// TIA Portal V17 export
// export: Created 2025-07-01T12:14:22.6243448Z, ExportSetting WithDefaults, DisplayName Totally Integrated Automation Portal, DisplayVersion V17, DisplayName TIA Portal Openness, DisplayVersion V17, DisplayName TIA Portal Version Control Interface, DisplayVersion V17, DisplayName SINAMICS Startdrive Advanced, DisplayVersion V17, DisplayName SINAMICS Startdrive G130, G150, S120, S150, SINAMICS MV, S210, DisplayVersion V17, DisplayName SINAMICS Startdrive G110M, G120, G120C, G120D, G120P, G115D, DisplayVersion V17, DisplayName STEP 7 Professional, DisplayVersion V17, DisplayName STEP 7 Safety, DisplayVersion V17, DisplayName WinCC Professional, DisplayVersion V17
FUNCTION_BLOCK "3PosLifter__Updated_V2_a4fa82_3a45ac7d-3c57-493c-83a9-58625a874be0 (3) - Copy_0df392"   // FB4, LAD
VERSION : 0.1
// stored: AutoNumber true, IsIECCheckEnabled false, UDAEnableTagReadback false
   VAR_INPUT
      L1S2Raise : Bool;
      iAreaClearConv : Bool;
      iAreaClearTransL2 : Bool;
      iAreaClear_TT : Bool;
      iAutoRunning : Bool;
      iErrorAck : Bool;
      iL1PalletPrsnt : Bool;
      iL1S1Raise : Bool;
      iL1S2Down : Bool;
      iL1S2DownOver : Bool;
      iL1S2Raise : Bool;
      iL2PalletPrsent : Bool;
      iL2S1Down : Bool;
      iL2S1Raise : Bool;
      iL2s2Raise : Bool;
      iLiffterAtPos1 : Bool;
      iLiffterAtPos2 : Bool;
      iLiffterAtPos3 : Bool;
      iLiffterAtPos4 : Bool;
      iLifterAt1 : Bool;
      iLifterAtPos1 : Bool;
      iLifterAtPos2 : Bool;
      iLifterAtPos3 : Bool;
      iLifterAtPos4 : Bool;
      iOTSFrmConv : Bool;
      iPalAtTT : Bool;
      iPalletAtL1 : Bool;
      iPalletAtL2 : Bool;
      iPalletAtLayre2 : Bool;
      iPalletAtTT : Bool;
      iPalletPrsntL1 : Bool;
      iRTRFrmConv : Bool;
      iRTRFrmTT : Bool;
      iRTRFrm_TT : Bool;
      iReacvAreaClr : Bool;
      iRecvAreaClear : Bool;
      iReset_fault : Bool;
      iRunOutActive : Bool;
      iRunOutCycle : Bool;
      iSstMode : Bool;
      iSstPB : Bool;
      iTransAreaClearConv : Bool;
      iTransAreaClr : Bool;
      ipalletPrsntAtTT : Bool;
   END_VAR
   VAR_OUTPUT
      qL1S1Down : Bool;
      qL1S1raise : Bool;
      qL1S2Down : Bool;
      qL1S2Raise : Bool;
      qL1TrnsfrConv : Bool;
      qL2S1raise : Bool;
      qL2S2Down : Bool;
      qL2S2Raise : Bool;
      qLiffterAtPos2 : Bool;
      qLifterAtPos1 : Bool;
      qLifterAtPos3 : Bool;
      qLifterAtPos4 : Bool;
      qLifterGotoPos1 : Bool;
      qOTSToNext : Bool;
      qOTSTo_TT : Bool;
      qOutput1 : Bool;
      qRTRToConv : Bool;
      qRTRToTT : Bool;
      qRTR_To_Conv : Bool;
   END_VAR
   VAR_IN_OUT
      IqRx_Frm_TT : Bool;
      iqRx_frm_Conv : Bool;
      iqTX_To_Conv : Bool;
      iqTX_To_TT : Bool;
      iqTx_To_ConvPos4 : Bool;
      iqTx_To_Rej : Bool;
   END_VAR
   VAR DB_SPECIFIC
      StateNo : Int;
      s100_StRunOutActive : Bool;
      s100_StRunOutActive_T1 : Bool;
      s100_StRunOutActive_T2 : Bool;
      s10_StRecovery : Bool;
      s10_StRecovery_T1 : Bool;
      s10_StRecovery_T2 : Bool;
      s10_StRecovery_T3 : Bool;
      s10_StRecovery_T4 : Bool;
      s10_StRecovery_T5 : Bool;
      s10_StRecovery_T6 : Bool;
      s10_StRecovery_T7 : Bool;
      s10_StRecovery_T8 : Bool;
      s110_InitialConvRun : Bool;
      s110_InitialConvRun_T1 : Bool;
      s120_StNextRdyInTransit : Bool;
      s120_StNextRdyInTransit_T1 : Bool;
      s120_StNextRdyInTransit_T2 : Bool;
      s130_StNextRdyInTransit_1 : Bool;
      s130_StNextRdyInTransit_1_T1 : Bool;
      s130_StNextRdyInTransit_1_T2 : Bool;
      s150_StWtLifterAtPosn1 : Bool;
      s150_StWtLifterAtPosn1_T1 : Bool;
      s15_StWtForFaultReset : Bool;
      s15_StWtForFaultReset_T1 : Bool;
      s160_StL1S2DownOver : Bool;
      s160_StL1S2DownOver_T1 : Bool;
      s170_StWtOTSFrmConv1 : Bool;
      s170_StWtOTSFrmConv1_T1 : Bool;
      s170_StWtOTSFrmConv1_T2 : Bool;
      s180_StWtRcvBegin : Bool;
      s180_StWtRcvBegin_T1 : Bool;
      s190_StWtL1RcvComplete : Bool;
      s190_StWtL1RcvComplete_T1 : Bool;
      s1_StWtResetRel : Bool;
      s1_StWtResetRel_T1 : Bool;
      s200_StWtForL1StprUp : Bool;
      s200_StWtForL1StprUp_T1 : Bool;
      s20_StWtForL1L2StoprsUp : Bool;
      s20_StWtForL1L2StoprsUp_T1 : Bool;
      s220_StWtL2S2Down : Bool;
      s220_StWtL2S2Down_T1 : Bool;
      s230_StWtL2TranBegin : Bool;
      s230_StWtL2TranBegin_T1 : Bool;
      s240_StWtL2TransComplete : Bool;
      s240_StWtL2TransComplete_T1 : Bool;
      s250_StWtDeforkDone : Bool;
      s250_StWtDeforkDone_Cond1 : Bool;
      s250_StWtDeforkDone_Cond2 : Bool;
      s250_StWtDeforkDone_T1 : Bool;
      s260_StChkRunOutActive1 : Bool;
      s260_StChkRunOutActive1_T1 : Bool;
      s260_StChkRunOutActive1_T2 : Bool;
      s270_StWtLifterAtPos4 : Bool;
      s270_StWtLifterAtPos4_T1 : Bool;
      s280_StWtRTRFrmConvPos4 : Bool;
      s280_StWtRTRFrmConvPos4_T1 : Bool;
      s285_StL1S2Down : Bool;
      s285_StL1S2Down_T1 : Bool;
      s290_StWtL1TransBeginPos4 : Bool;
      s290_StWtL1TransBeginPos4_T1 : Bool;
      s300_StWtTransDonePos4 : Bool;
      s300_StWtTransDonePos4_T1 : Bool;
      s30_StChkPalletPrsntL1L2 : Bool;
      s30_StChkPalletPrsntL1L2_T1 : Bool;
      s30_StChkPalletPrsntL1L2_T2 : Bool;
      s30_StChkPalletPrsntL1L2_T3 : Bool;
      s30_StChkPalletPrsntL1L2_T4 : Bool;
      s310_StChkPalletAtTT1 : Bool;
      s310_StChkPalletAtTT1_T1 : Bool;
      s310_StChkPalletAtTT1_T2 : Bool;
      s320_StWtLifterAtPos3 : Bool;
      s320_StWtLifterAtPos3_T1 : Bool;
      s330_StWtL2S1Down : Bool;
      s330_StWtL2S1Down_T1 : Bool;
      s340_StWtOTSFrmTT : Bool;
      s340_StWtOTSFrmTT_T1 : Bool;
      s350_StWtL2RecvingActive : Bool;
      s350_StWtL2RecvingActive_T1 : Bool;
      s360_StWtL2RcvDone : Bool;
      s360_StWtL2RcvDone_T1 : Bool;
      s370_StChkPalAtTT : Bool;
      s370_StChkPalAtTT_T1 : Bool;
      s370_StChkPalAtTT_T2 : Bool;
      s370_StChkPalAtTT_T3 : Bool;
      s380_StWtLifterAtPos2 : Bool;
      s380_StWtLifterAtPos2_T1 : Bool;
      s390_StWtRTRFrmTT : Bool;
      s390_StWtRTRFrmTT_T1 : Bool;
      s400_StWtL1S1Down1 : Bool;
      s400_StWtL1S1Down1_T1 : Bool;
      s40_StChkPalletAtTT : Bool;
      s40_StChkPalletAtTT_T1 : Bool;
      s40_StChkPalletAtTT_T2 : Bool;
      s410_StWtL1TransBegin : Bool;
      s410_StWtL1TransBegin_T1 : Bool;
      s420_StWtL1TransComplet : Bool;
      s420_StWtL1TransComplet_T1 : Bool;
      s430_StNextRdyInTransit_3 : Bool;
      s430_StNextRdyInTransit_3_T1 : Bool;
      s430_StNextRdyInTransit_3_T2 : Bool;
      s50_StWtLifterAtPos1 : Bool;
      s50_StWtLifterAtPos1_T1 : Bool;
      s60_StWtL1S2DownOver : Bool;
      s60_StWtL1S2DownOver_T1 : Bool;
      s70_StWtOTSFrmConv : Bool;
      s70_StWtOTSFrmConv_T1 : Bool;
      s80_StWtL1RecvBegin : Bool;
      s80_StWtL1RecvBegin_T1 : Bool;
      s90_StWtL1PalRcvDone : Bool;
      s90_StWtL1PalRcvDone_T1 : Bool;
      sOTSTimeout : Struct
         q : Bool;
      END_STRUCT;
      sSeq1Over : Bool;
      sSeq2Over : Bool;
      sSst : Bool;
      sSstPulse : Bool;
      sSstRise : Bool;
      sStWtResetRel : Bool;
      sStWtResetRel_T1 : Bool;
   END_VAR
   VAR_TEMP
      tOne : Bool;
   END_VAR
   VAR_TEMP   // added for the SCL form of the ladder/FBD networks
      _w1 : Bool;
   END_VAR
BEGIN

REGION Network 1
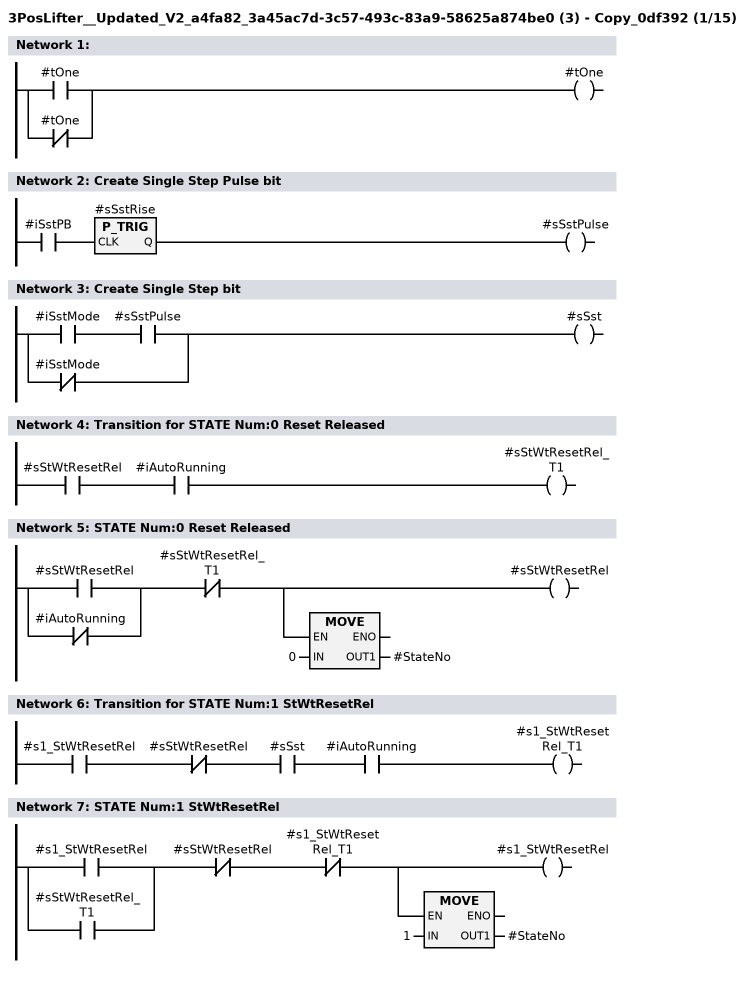
   RUNG wire#powerrail
      Contact( #tOne )
      wire#w1
      Coil( #tOne )
   END_RUNG
   RUNG wire#powerrail
      I_Contact( #tOne )
   END_RUNG wire#w1
   // the same network as SCL:
   #tOne := #tOne OR NOT #tOne;
END_REGION

REGION Network 2: Create Single Step Pulse bit
   RUNG wire#powerrail
      Contact( #iSstPB )
      P_Trig( #sSstRise )
      Coil( #sSstPulse )
   END_RUNG
   // the same network as SCL:
   #_w1 := #iSstPB AND NOT #sSstRise;   // rising edge
   #sSstRise := #iSstPB;
   #sSstPulse := #_w1;
END_REGION

REGION Network 3: Create Single Step bit
   RUNG wire#powerrail
      Contact( #iSstMode )
      Contact( #sSstPulse )
      wire#w1
      Coil( #sSst )
   END_RUNG
   RUNG wire#powerrail
      I_Contact( #iSstMode )
   END_RUNG wire#w1
   // the same network as SCL:
   #sSst := (#iSstMode AND #sSstPulse) OR NOT #iSstMode;
END_REGION

REGION Network 4: Transition for STATE Num:0 Reset Released
   RUNG wire#powerrail
      Contact( #sStWtResetRel )
      Contact( #iAutoRunning )
      Coil( #sStWtResetRel_T1 )
   END_RUNG
   // the same network as SCL:
   #sStWtResetRel_T1 := #sStWtResetRel AND #iAutoRunning;
END_REGION

REGION Network 5: STATE Num:0 Reset Released
   RUNG wire#powerrail
      Contact( #sStWtResetRel )
      wire#w1
      I_Contact( #sStWtResetRel_T1 )
      wire#w2
      Coil( #sStWtResetRel )
   END_RUNG
   RUNG wire#powerrail
      I_Contact( #iAutoRunning )
   END_RUNG wire#w1
   RUNG wire#w2
      { S7_GenerateENO := "TRUE" } Move(in := 0, out1 => #StateNo)
   END_RUNG
   // the same network as SCL:
   #sStWtResetRel := (#sStWtResetRel OR NOT #iAutoRunning) AND NOT #sStWtResetRel_T1;
   IF #sStWtResetRel THEN #StateNo := 0; END_IF;
END_REGION

REGION Network 6: Transition for STATE Num:1 StWtResetRel
   RUNG wire#powerrail
      Contact( #s1_StWtResetRel )
      I_Contact( #sStWtResetRel )
      Contact( #sSst )
      Contact( #iAutoRunning )
      Coil( #s1_StWtResetRel_T1 )
   END_RUNG
   // the same network as SCL:
   #s1_StWtResetRel_T1 := #s1_StWtResetRel AND NOT #sStWtResetRel AND #sSst AND #iAutoRunning;
END_REGION

REGION Network 7: STATE Num:1 StWtResetRel
   RUNG wire#powerrail
      Contact( #s1_StWtResetRel )
      wire#w1
      I_Contact( #sStWtResetRel )
      I_Contact( #s1_StWtResetRel_T1 )
      wire#w2
      Coil( #s1_StWtResetRel )
   END_RUNG
   RUNG wire#powerrail
      Contact( #sStWtResetRel_T1 )
   END_RUNG wire#w1
   RUNG wire#w2
      { S7_GenerateENO := "TRUE" } Move(in := 1, out1 => #StateNo)
   END_RUNG
   // the same network as SCL:
   #s1_StWtResetRel := (#s1_StWtResetRel OR #sStWtResetRel_T1) AND NOT #sStWtResetRel AND NOT #s1_StWtResetRel_T1;
   IF #s1_StWtResetRel THEN #StateNo := 1; END_IF;
END_REGION

REGION Network 8: Transition for STATE Num:10 StRecovery
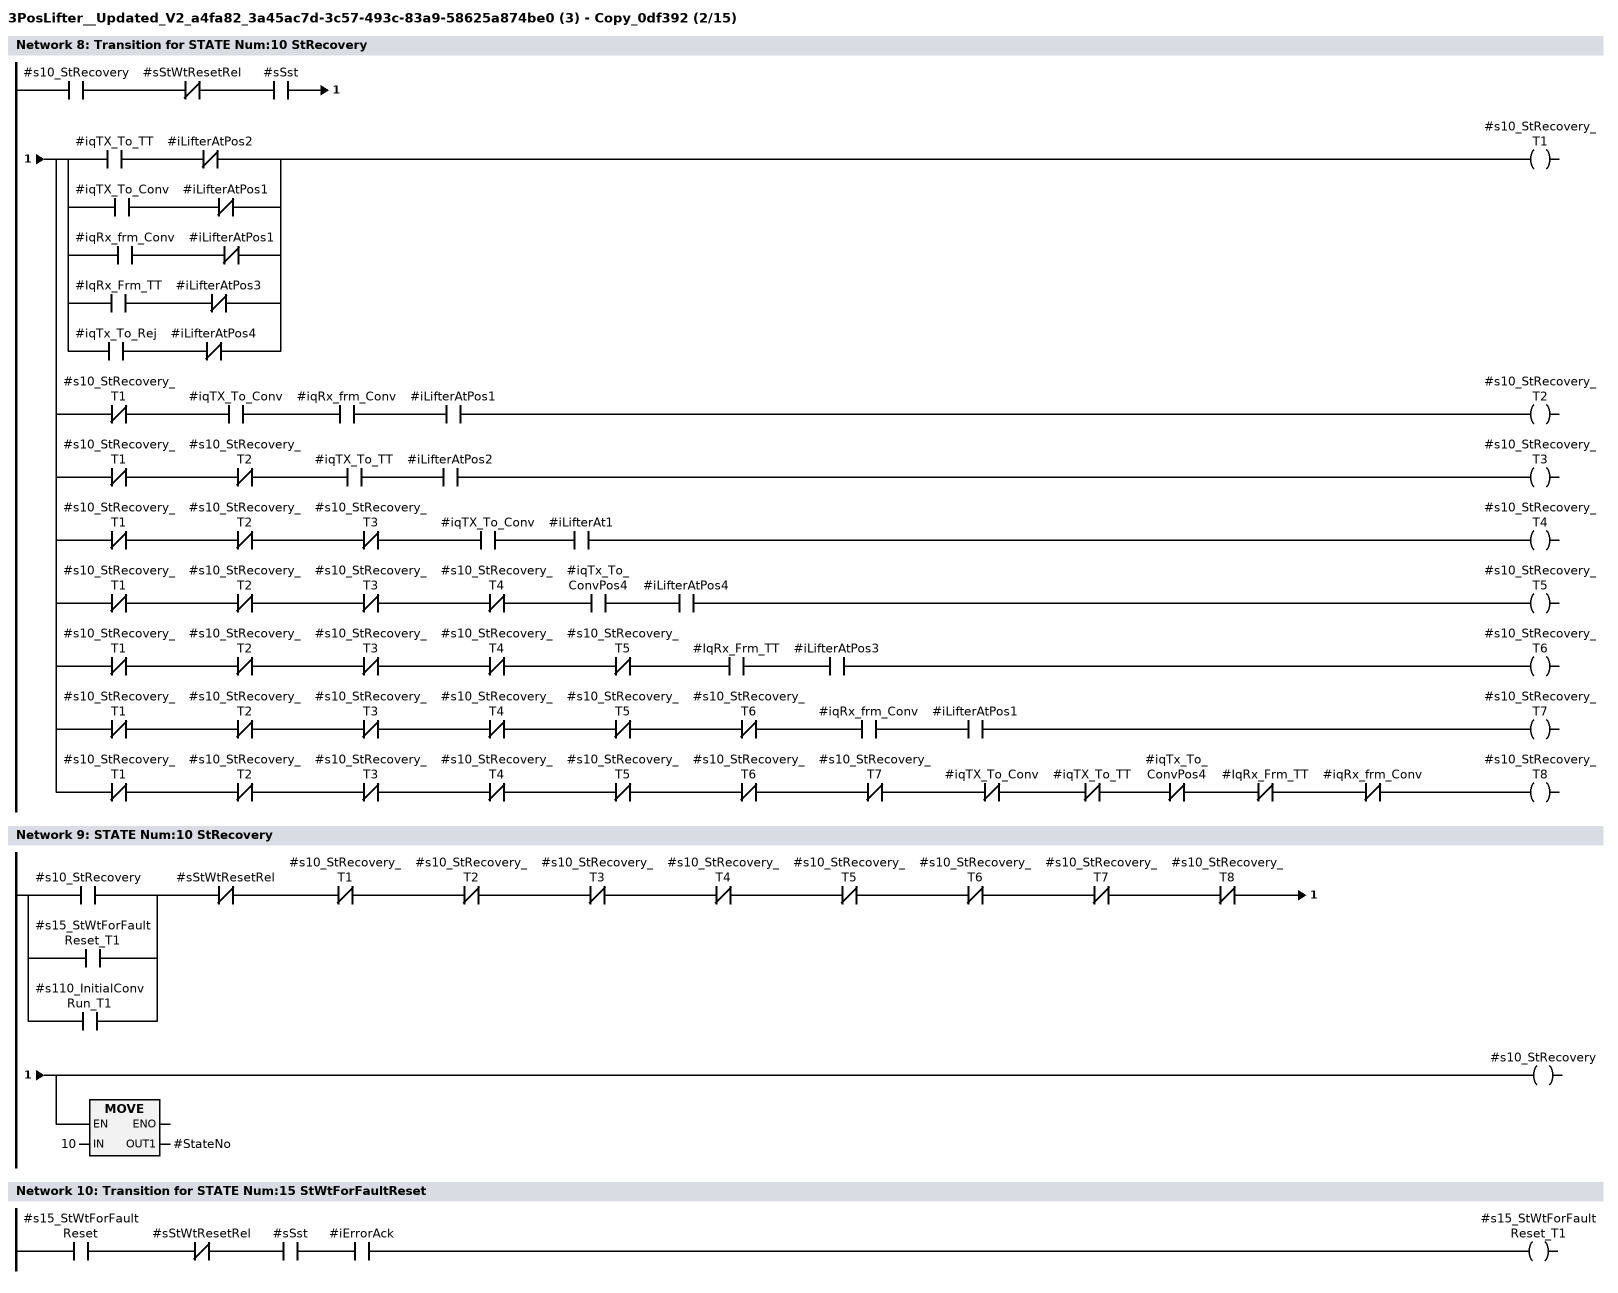
   RUNG wire#powerrail
      Contact( #s10_StRecovery )
      I_Contact( #sStWtResetRel )
      Contact( #sSst )
      wire#w1
      Contact( #iqTX_To_TT )
      I_Contact( #iLifterAtPos2 )
      wire#w2
      Coil( #s10_StRecovery_T1 )
   END_RUNG
   RUNG wire#w1
      Contact( #iqTX_To_Conv )
      I_Contact( #iLifterAtPos1 )
   END_RUNG wire#w2
   RUNG wire#w1
      Contact( #iqRx_frm_Conv )
      I_Contact( #iLifterAtPos1 )
   END_RUNG wire#w2
   RUNG wire#w1
      Contact( #IqRx_Frm_TT )
      I_Contact( #iLifterAtPos3 )
   END_RUNG wire#w2
   RUNG wire#w1
      Contact( #iqTx_To_Rej )
      I_Contact( #iLifterAtPos4 )
   END_RUNG wire#w2
   RUNG wire#w1
      I_Contact( #s10_StRecovery_T1 )
      Contact( #iqTX_To_Conv )
      Contact( #iqRx_frm_Conv )
      Contact( #iLifterAtPos1 )
      Coil( #s10_StRecovery_T2 )
   END_RUNG
   RUNG wire#w1
      I_Contact( #s10_StRecovery_T1 )
      I_Contact( #s10_StRecovery_T2 )
      Contact( #iqTX_To_TT )
      Contact( #iLifterAtPos2 )
      Coil( #s10_StRecovery_T3 )
   END_RUNG
   RUNG wire#w1
      I_Contact( #s10_StRecovery_T1 )
      I_Contact( #s10_StRecovery_T2 )
      I_Contact( #s10_StRecovery_T3 )
      Contact( #iqTX_To_Conv )
      Contact( #iLifterAt1 )
      Coil( #s10_StRecovery_T4 )
   END_RUNG
   RUNG wire#w1
      I_Contact( #s10_StRecovery_T1 )
      I_Contact( #s10_StRecovery_T2 )
      I_Contact( #s10_StRecovery_T3 )
      I_Contact( #s10_StRecovery_T4 )
      Contact( #iqTx_To_ConvPos4 )
      Contact( #iLifterAtPos4 )
      Coil( #s10_StRecovery_T5 )
   END_RUNG
   RUNG wire#w1
      I_Contact( #s10_StRecovery_T1 )
      I_Contact( #s10_StRecovery_T2 )
      I_Contact( #s10_StRecovery_T3 )
      I_Contact( #s10_StRecovery_T4 )
      I_Contact( #s10_StRecovery_T5 )
      Contact( #IqRx_Frm_TT )
      Contact( #iLifterAtPos3 )
      Coil( #s10_StRecovery_T6 )
   END_RUNG
   RUNG wire#w1
      I_Contact( #s10_StRecovery_T1 )
      I_Contact( #s10_StRecovery_T2 )
      I_Contact( #s10_StRecovery_T3 )
      I_Contact( #s10_StRecovery_T4 )
      I_Contact( #s10_StRecovery_T5 )
      I_Contact( #s10_StRecovery_T6 )
      Contact( #iqRx_frm_Conv )
      Contact( #iLifterAtPos1 )
      Coil( #s10_StRecovery_T7 )
   END_RUNG
   RUNG wire#w1
      I_Contact( #s10_StRecovery_T1 )
      I_Contact( #s10_StRecovery_T2 )
      I_Contact( #s10_StRecovery_T3 )
      I_Contact( #s10_StRecovery_T4 )
      I_Contact( #s10_StRecovery_T5 )
      I_Contact( #s10_StRecovery_T6 )
      I_Contact( #s10_StRecovery_T7 )
      I_Contact( #iqTX_To_Conv )
      I_Contact( #iqTX_To_TT )
      I_Contact( #iqTx_To_ConvPos4 )
      I_Contact( #IqRx_Frm_TT )
      I_Contact( #iqRx_frm_Conv )
      Coil( #s10_StRecovery_T8 )
   END_RUNG
   // the same network as SCL:
   #_w1 := #s10_StRecovery AND NOT #sStWtResetRel AND #sSst;
   #s10_StRecovery_T1 := #_w1 AND ((#iqTX_To_TT AND NOT #iLifterAtPos2) OR (#iqTX_To_Conv AND NOT #iLifterAtPos1) OR (#iqRx_frm_Conv AND NOT #iLifterAtPos1) OR (#IqRx_Frm_TT AND NOT #iLifterAtPos3) OR (#iqTx_To_Rej AND NOT #iLifterAtPos4));
   #s10_StRecovery_T2 := #_w1 AND NOT #s10_StRecovery_T1 AND #iqTX_To_Conv AND #iqRx_frm_Conv AND #iLifterAtPos1;
   #s10_StRecovery_T3 := #_w1 AND NOT #s10_StRecovery_T1 AND NOT #s10_StRecovery_T2 AND #iqTX_To_TT AND #iLifterAtPos2;
   #s10_StRecovery_T4 := #_w1 AND NOT #s10_StRecovery_T1 AND NOT #s10_StRecovery_T2 AND NOT #s10_StRecovery_T3 AND #iqTX_To_Conv AND #iLifterAt1;
   #s10_StRecovery_T5 := #_w1 AND NOT #s10_StRecovery_T1 AND NOT #s10_StRecovery_T2 AND NOT #s10_StRecovery_T3 AND NOT #s10_StRecovery_T4 AND #iqTx_To_ConvPos4 AND #iLifterAtPos4;
   #s10_StRecovery_T6 := #_w1 AND NOT #s10_StRecovery_T1 AND NOT #s10_StRecovery_T2 AND NOT #s10_StRecovery_T3 AND NOT #s10_StRecovery_T4 AND NOT #s10_StRecovery_T5 AND #IqRx_Frm_TT AND #iLifterAtPos3;
   #s10_StRecovery_T7 := #_w1 AND NOT #s10_StRecovery_T1 AND NOT #s10_StRecovery_T2 AND NOT #s10_StRecovery_T3 AND NOT #s10_StRecovery_T4 AND NOT #s10_StRecovery_T5 AND NOT #s10_StRecovery_T6 AND #iqRx_frm_Conv AND #iLifterAtPos1;
   #s10_StRecovery_T8 := #_w1 AND NOT #s10_StRecovery_T1 AND NOT #s10_StRecovery_T2 AND NOT #s10_StRecovery_T3 AND NOT #s10_StRecovery_T4 AND NOT #s10_StRecovery_T5 AND NOT #s10_StRecovery_T6 AND NOT #s10_StRecovery_T7 AND NOT #iqTX_To_Conv AND NOT #iqTX_To_TT AND NOT #iqTx_To_ConvPos4 AND NOT #IqRx_Frm_TT AND NOT #iqRx_frm_Conv;
END_REGION

REGION Network 9: STATE Num:10 StRecovery
   RUNG wire#powerrail
      Contact( #s10_StRecovery )
      wire#w1
      I_Contact( #sStWtResetRel )
      I_Contact( #s10_StRecovery_T1 )
      I_Contact( #s10_StRecovery_T2 )
      I_Contact( #s10_StRecovery_T3 )
      I_Contact( #s10_StRecovery_T4 )
      I_Contact( #s10_StRecovery_T5 )
      I_Contact( #s10_StRecovery_T6 )
      I_Contact( #s10_StRecovery_T7 )
      I_Contact( #s10_StRecovery_T8 )
      wire#w2
      Coil( #s10_StRecovery )
   END_RUNG
   RUNG wire#powerrail
      Contact( #s15_StWtForFaultReset_T1 )
   END_RUNG wire#w1
   RUNG wire#powerrail
      Contact( #s110_InitialConvRun_T1 )
   END_RUNG wire#w1
   RUNG wire#w2
      { S7_GenerateENO := "TRUE" } Move(in := 10, out1 => #StateNo)
   END_RUNG
   // the same network as SCL:
   #s10_StRecovery := (#s10_StRecovery OR #s15_StWtForFaultReset_T1 OR #s110_InitialConvRun_T1) AND NOT #sStWtResetRel AND NOT #s10_StRecovery_T1 AND NOT #s10_StRecovery_T2 AND NOT #s10_StRecovery_T3 AND NOT #s10_StRecovery_T4 AND NOT #s10_StRecovery_T5 AND NOT #s10_StRecovery_T6 AND NOT #s10_StRecovery_T7 AND NOT #s10_StRecovery_T8;
   IF #s10_StRecovery THEN #StateNo := 10; END_IF;
END_REGION

REGION Network 10: Transition for STATE Num:15 StWtForFaultReset
   RUNG wire#powerrail
      Contact( #s15_StWtForFaultReset )
      I_Contact( #sStWtResetRel )
      Contact( #sSst )
      Contact( #iErrorAck )
      Coil( #s15_StWtForFaultReset_T1 )
   END_RUNG
   // the same network as SCL:
   #s15_StWtForFaultReset_T1 := #s15_StWtForFaultReset AND NOT #sStWtResetRel AND #sSst AND #iErrorAck;
END_REGION

REGION Network 11: STATE Num:15 StWtForFaultReset
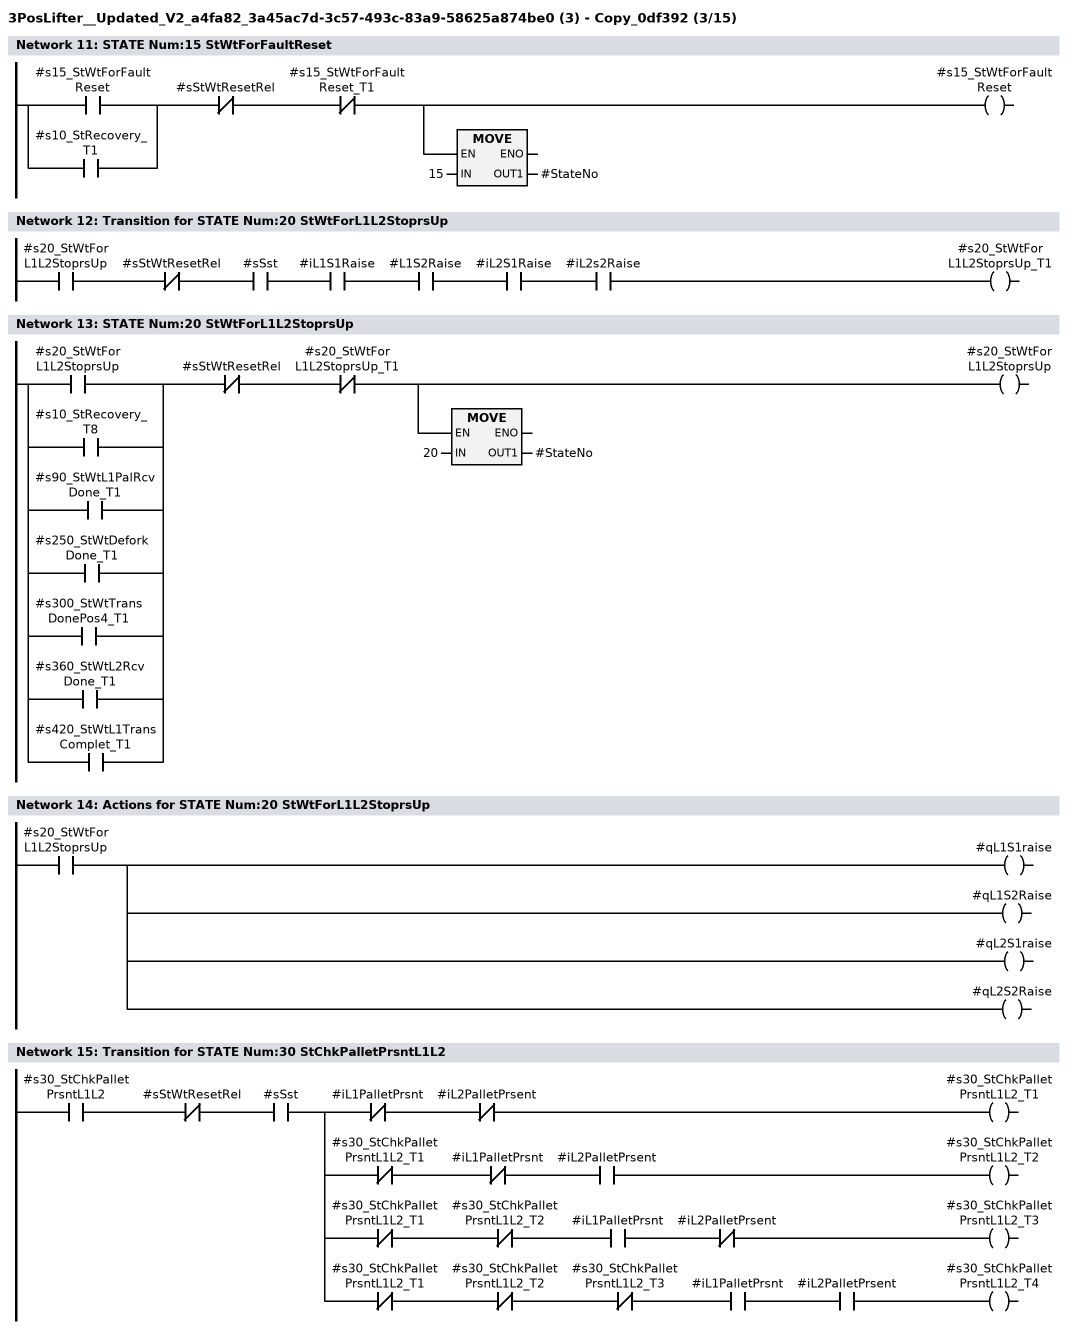
   RUNG wire#powerrail
      Contact( #s15_StWtForFaultReset )
      wire#w1
      I_Contact( #sStWtResetRel )
      I_Contact( #s15_StWtForFaultReset_T1 )
      wire#w2
      Coil( #s15_StWtForFaultReset )
   END_RUNG
   RUNG wire#powerrail
      Contact( #s10_StRecovery_T1 )
   END_RUNG wire#w1
   RUNG wire#w2
      { S7_GenerateENO := "TRUE" } Move(in := 15, out1 => #StateNo)
   END_RUNG
   // the same network as SCL:
   #s15_StWtForFaultReset := (#s15_StWtForFaultReset OR #s10_StRecovery_T1) AND NOT #sStWtResetRel AND NOT #s15_StWtForFaultReset_T1;
   IF #s15_StWtForFaultReset THEN #StateNo := 15; END_IF;
END_REGION

REGION Network 12: Transition for STATE Num:20 StWtForL1L2StoprsUp
   RUNG wire#powerrail
      Contact( #s20_StWtForL1L2StoprsUp )
      I_Contact( #sStWtResetRel )
      Contact( #sSst )
      Contact( #iL1S1Raise )
      Contact( #L1S2Raise )
      Contact( #iL2S1Raise )
      Contact( #iL2s2Raise )
      Coil( #s20_StWtForL1L2StoprsUp_T1 )
   END_RUNG
   // the same network as SCL:
   #s20_StWtForL1L2StoprsUp_T1 := #s20_StWtForL1L2StoprsUp AND NOT #sStWtResetRel AND #sSst AND #iL1S1Raise AND #L1S2Raise AND #iL2S1Raise AND #iL2s2Raise;
END_REGION

REGION Network 13: STATE Num:20 StWtForL1L2StoprsUp
   RUNG wire#powerrail
      Contact( #s20_StWtForL1L2StoprsUp )
      wire#w1
      I_Contact( #sStWtResetRel )
      I_Contact( #s20_StWtForL1L2StoprsUp_T1 )
      wire#w2
      Coil( #s20_StWtForL1L2StoprsUp )
   END_RUNG
   RUNG wire#powerrail
      Contact( #s10_StRecovery_T8 )
   END_RUNG wire#w1
   RUNG wire#powerrail
      Contact( #s90_StWtL1PalRcvDone_T1 )
   END_RUNG wire#w1
   RUNG wire#powerrail
      Contact( #s250_StWtDeforkDone_T1 )
   END_RUNG wire#w1
   RUNG wire#powerrail
      Contact( #s300_StWtTransDonePos4_T1 )
   END_RUNG wire#w1
   RUNG wire#powerrail
      Contact( #s360_StWtL2RcvDone_T1 )
   END_RUNG wire#w1
   RUNG wire#powerrail
      Contact( #s420_StWtL1TransComplet_T1 )
   END_RUNG wire#w1
   RUNG wire#w2
      { S7_GenerateENO := "TRUE" } Move(in := 20, out1 => #StateNo)
   END_RUNG
   // the same network as SCL:
   #s20_StWtForL1L2StoprsUp := (#s20_StWtForL1L2StoprsUp OR #s10_StRecovery_T8 OR #s90_StWtL1PalRcvDone_T1 OR #s250_StWtDeforkDone_T1 OR #s300_StWtTransDonePos4_T1 OR #s360_StWtL2RcvDone_T1 OR #s420_StWtL1TransComplet_T1) AND NOT #sStWtResetRel AND NOT #s20_StWtForL1L2StoprsUp_T1;
   IF #s20_StWtForL1L2StoprsUp THEN #StateNo := 20; END_IF;
END_REGION

REGION Network 14: Actions for STATE Num:20 StWtForL1L2StoprsUp
   RUNG wire#powerrail
      Contact( #s20_StWtForL1L2StoprsUp )
      wire#w1
      Coil( #qL1S1raise )
   END_RUNG
   RUNG wire#w1
      Coil( #qL1S2Raise )
   END_RUNG
   RUNG wire#w1
      Coil( #qL2S1raise )
   END_RUNG
   RUNG wire#w1
      Coil( #qL2S2Raise )
   END_RUNG
   // the same network as SCL:
   #qL1S1raise := #s20_StWtForL1L2StoprsUp;
   #qL1S2Raise := #s20_StWtForL1L2StoprsUp;
   #qL2S1raise := #s20_StWtForL1L2StoprsUp;
   #qL2S2Raise := #s20_StWtForL1L2StoprsUp;
END_REGION

REGION Network 15: Transition for STATE Num:30 StChkPalletPrsntL1L2
   RUNG wire#powerrail
      Contact( #s30_StChkPalletPrsntL1L2 )
      I_Contact( #sStWtResetRel )
      Contact( #sSst )
      wire#w1
      I_Contact( #iL1PalletPrsnt )
      I_Contact( #iL2PalletPrsent )
      Coil( #s30_StChkPalletPrsntL1L2_T1 )
   END_RUNG
   RUNG wire#w1
      I_Contact( #s30_StChkPalletPrsntL1L2_T1 )
      I_Contact( #iL1PalletPrsnt )
      Contact( #iL2PalletPrsent )
      Coil( #s30_StChkPalletPrsntL1L2_T2 )
   END_RUNG
   RUNG wire#w1
      I_Contact( #s30_StChkPalletPrsntL1L2_T1 )
      I_Contact( #s30_StChkPalletPrsntL1L2_T2 )
      Contact( #iL1PalletPrsnt )
      I_Contact( #iL2PalletPrsent )
      Coil( #s30_StChkPalletPrsntL1L2_T3 )
   END_RUNG
   RUNG wire#w1
      I_Contact( #s30_StChkPalletPrsntL1L2_T1 )
      I_Contact( #s30_StChkPalletPrsntL1L2_T2 )
      I_Contact( #s30_StChkPalletPrsntL1L2_T3 )
      Contact( #iL1PalletPrsnt )
      Contact( #iL2PalletPrsent )
      Coil( #s30_StChkPalletPrsntL1L2_T4 )
   END_RUNG
   // the same network as SCL:
   #_w1 := #s30_StChkPalletPrsntL1L2 AND NOT #sStWtResetRel AND #sSst;
   #s30_StChkPalletPrsntL1L2_T1 := #_w1 AND NOT #iL1PalletPrsnt AND NOT #iL2PalletPrsent;
   #s30_StChkPalletPrsntL1L2_T2 := #_w1 AND NOT #s30_StChkPalletPrsntL1L2_T1 AND NOT #iL1PalletPrsnt AND #iL2PalletPrsent;
   #s30_StChkPalletPrsntL1L2_T3 := #_w1 AND NOT #s30_StChkPalletPrsntL1L2_T1 AND NOT #s30_StChkPalletPrsntL1L2_T2 AND #iL1PalletPrsnt AND NOT #iL2PalletPrsent;
   #s30_StChkPalletPrsntL1L2_T4 := #_w1 AND NOT #s30_StChkPalletPrsntL1L2_T1 AND NOT #s30_StChkPalletPrsntL1L2_T2 AND NOT #s30_StChkPalletPrsntL1L2_T3 AND #iL1PalletPrsnt AND #iL2PalletPrsent;
END_REGION

REGION Network 16: STATE Num:30 StChkPalletPrsntL1L2
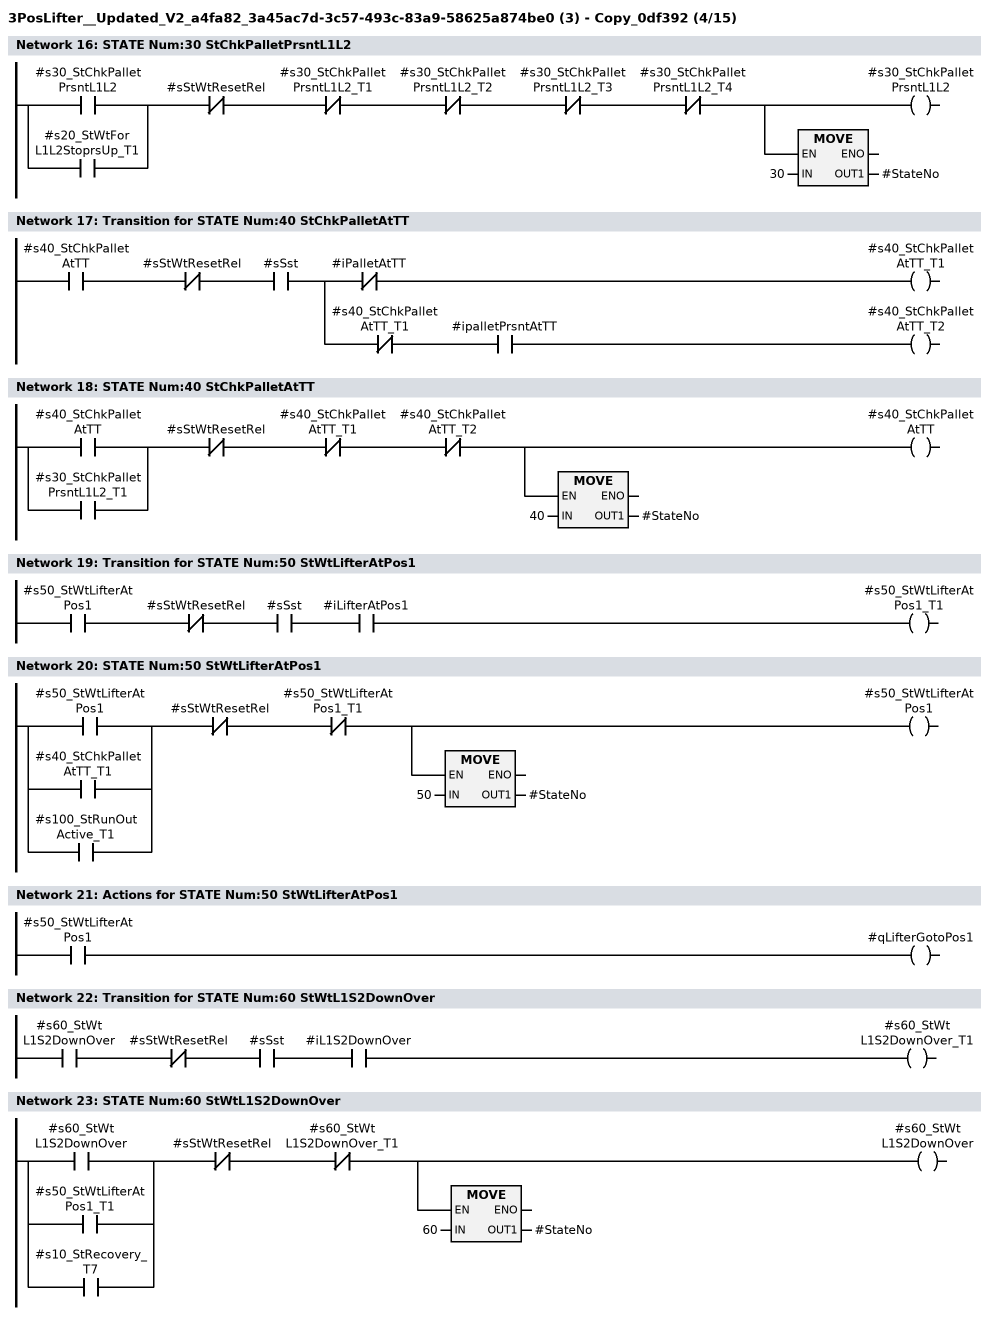
   RUNG wire#powerrail
      Contact( #s30_StChkPalletPrsntL1L2 )
      wire#w1
      I_Contact( #sStWtResetRel )
      I_Contact( #s30_StChkPalletPrsntL1L2_T1 )
      I_Contact( #s30_StChkPalletPrsntL1L2_T2 )
      I_Contact( #s30_StChkPalletPrsntL1L2_T3 )
      I_Contact( #s30_StChkPalletPrsntL1L2_T4 )
      wire#w2
      Coil( #s30_StChkPalletPrsntL1L2 )
   END_RUNG
   RUNG wire#powerrail
      Contact( #s20_StWtForL1L2StoprsUp_T1 )
   END_RUNG wire#w1
   RUNG wire#w2
      { S7_GenerateENO := "TRUE" } Move(in := 30, out1 => #StateNo)
   END_RUNG
   // the same network as SCL:
   #s30_StChkPalletPrsntL1L2 := (#s30_StChkPalletPrsntL1L2 OR #s20_StWtForL1L2StoprsUp_T1) AND NOT #sStWtResetRel AND NOT #s30_StChkPalletPrsntL1L2_T1 AND NOT #s30_StChkPalletPrsntL1L2_T2 AND NOT #s30_StChkPalletPrsntL1L2_T3 AND NOT #s30_StChkPalletPrsntL1L2_T4;
   IF #s30_StChkPalletPrsntL1L2 THEN #StateNo := 30; END_IF;
END_REGION

REGION Network 17: Transition for STATE Num:40 StChkPalletAtTT
   RUNG wire#powerrail
      Contact( #s40_StChkPalletAtTT )
      I_Contact( #sStWtResetRel )
      Contact( #sSst )
      wire#w1
      I_Contact( #iPalletAtTT )
      Coil( #s40_StChkPalletAtTT_T1 )
   END_RUNG
   RUNG wire#w1
      I_Contact( #s40_StChkPalletAtTT_T1 )
      Contact( #ipalletPrsntAtTT )
      Coil( #s40_StChkPalletAtTT_T2 )
   END_RUNG
   // the same network as SCL:
   #_w1 := #s40_StChkPalletAtTT AND NOT #sStWtResetRel AND #sSst;
   #s40_StChkPalletAtTT_T1 := #_w1 AND NOT #iPalletAtTT;
   #s40_StChkPalletAtTT_T2 := #_w1 AND NOT #s40_StChkPalletAtTT_T1 AND #ipalletPrsntAtTT;
END_REGION

REGION Network 18: STATE Num:40 StChkPalletAtTT
   RUNG wire#powerrail
      Contact( #s40_StChkPalletAtTT )
      wire#w1
      I_Contact( #sStWtResetRel )
      I_Contact( #s40_StChkPalletAtTT_T1 )
      I_Contact( #s40_StChkPalletAtTT_T2 )
      wire#w2
      Coil( #s40_StChkPalletAtTT )
   END_RUNG
   RUNG wire#powerrail
      Contact( #s30_StChkPalletPrsntL1L2_T1 )
   END_RUNG wire#w1
   RUNG wire#w2
      { S7_GenerateENO := "TRUE" } Move(in := 40, out1 => #StateNo)
   END_RUNG
   // the same network as SCL:
   #s40_StChkPalletAtTT := (#s40_StChkPalletAtTT OR #s30_StChkPalletPrsntL1L2_T1) AND NOT #sStWtResetRel AND NOT #s40_StChkPalletAtTT_T1 AND NOT #s40_StChkPalletAtTT_T2;
   IF #s40_StChkPalletAtTT THEN #StateNo := 40; END_IF;
END_REGION

REGION Network 19: Transition for STATE Num:50 StWtLifterAtPos1
   RUNG wire#powerrail
      Contact( #s50_StWtLifterAtPos1 )
      I_Contact( #sStWtResetRel )
      Contact( #sSst )
      Contact( #iLifterAtPos1 )
      Coil( #s50_StWtLifterAtPos1_T1 )
   END_RUNG
   // the same network as SCL:
   #s50_StWtLifterAtPos1_T1 := #s50_StWtLifterAtPos1 AND NOT #sStWtResetRel AND #sSst AND #iLifterAtPos1;
END_REGION

REGION Network 20: STATE Num:50 StWtLifterAtPos1
   RUNG wire#powerrail
      Contact( #s50_StWtLifterAtPos1 )
      wire#w1
      I_Contact( #sStWtResetRel )
      I_Contact( #s50_StWtLifterAtPos1_T1 )
      wire#w2
      Coil( #s50_StWtLifterAtPos1 )
   END_RUNG
   RUNG wire#powerrail
      Contact( #s40_StChkPalletAtTT_T1 )
   END_RUNG wire#w1
   RUNG wire#powerrail
      Contact( #s100_StRunOutActive_T1 )
   END_RUNG wire#w1
   RUNG wire#w2
      { S7_GenerateENO := "TRUE" } Move(in := 50, out1 => #StateNo)
   END_RUNG
   // the same network as SCL:
   #s50_StWtLifterAtPos1 := (#s50_StWtLifterAtPos1 OR #s40_StChkPalletAtTT_T1 OR #s100_StRunOutActive_T1) AND NOT #sStWtResetRel AND NOT #s50_StWtLifterAtPos1_T1;
   IF #s50_StWtLifterAtPos1 THEN #StateNo := 50; END_IF;
END_REGION

REGION Network 21: Actions for STATE Num:50 StWtLifterAtPos1
   RUNG wire#powerrail
      Contact( #s50_StWtLifterAtPos1 )
      Coil( #qLifterGotoPos1 )
   END_RUNG
   // the same network as SCL:
   #qLifterGotoPos1 := #s50_StWtLifterAtPos1;
END_REGION

REGION Network 22: Transition for STATE Num:60 StWtL1S2DownOver
   RUNG wire#powerrail
      Contact( #s60_StWtL1S2DownOver )
      I_Contact( #sStWtResetRel )
      Contact( #sSst )
      Contact( #iL1S2DownOver )
      Coil( #s60_StWtL1S2DownOver_T1 )
   END_RUNG
   // the same network as SCL:
   #s60_StWtL1S2DownOver_T1 := #s60_StWtL1S2DownOver AND NOT #sStWtResetRel AND #sSst AND #iL1S2DownOver;
END_REGION

REGION Network 23: STATE Num:60 StWtL1S2DownOver
   RUNG wire#powerrail
      Contact( #s60_StWtL1S2DownOver )
      wire#w1
      I_Contact( #sStWtResetRel )
      I_Contact( #s60_StWtL1S2DownOver_T1 )
      wire#w2
      Coil( #s60_StWtL1S2DownOver )
   END_RUNG
   RUNG wire#powerrail
      Contact( #s50_StWtLifterAtPos1_T1 )
   END_RUNG wire#w1
   RUNG wire#powerrail
      Contact( #s10_StRecovery_T7 )
   END_RUNG wire#w1
   RUNG wire#w2
      { S7_GenerateENO := "TRUE" } Move(in := 60, out1 => #StateNo)
   END_RUNG
   // the same network as SCL:
   #s60_StWtL1S2DownOver := (#s60_StWtL1S2DownOver OR #s50_StWtLifterAtPos1_T1 OR #s10_StRecovery_T7) AND NOT #sStWtResetRel AND NOT #s60_StWtL1S2DownOver_T1;
   IF #s60_StWtL1S2DownOver THEN #StateNo := 60; END_IF;
END_REGION

REGION Network 24: Actions for STATE Num:60 StWtL1S2DownOver
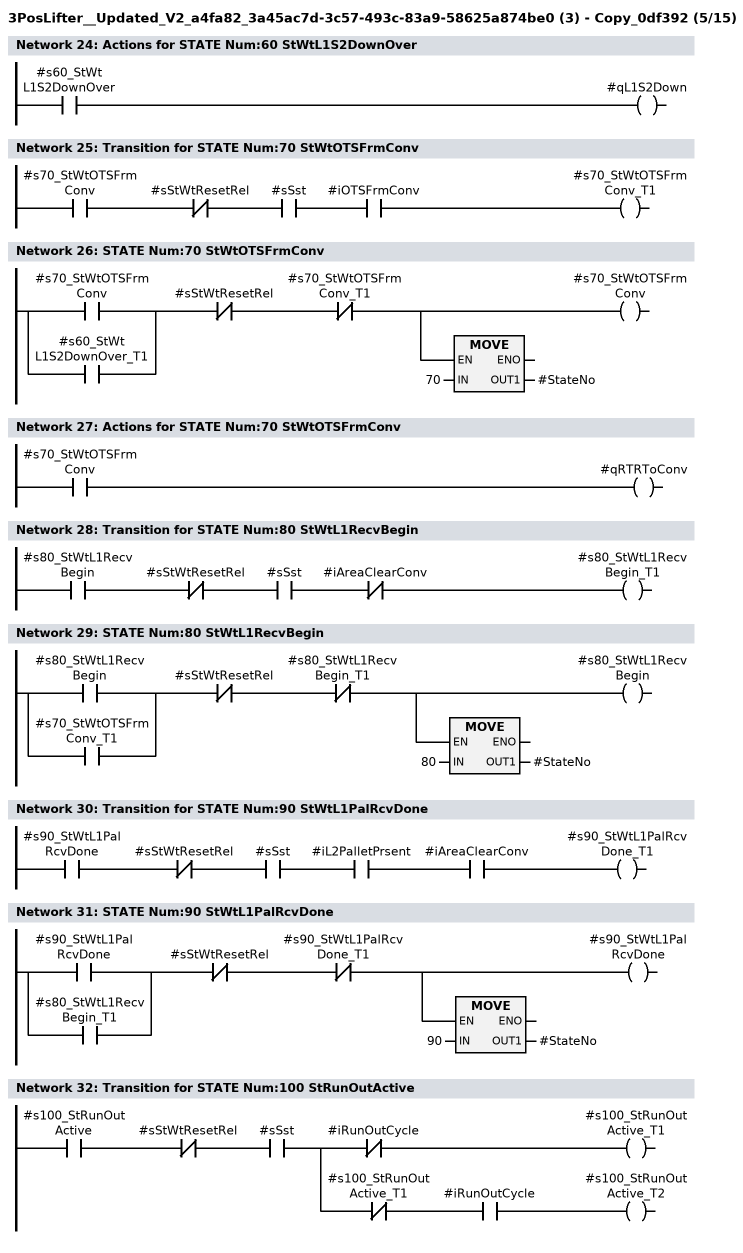
   RUNG wire#powerrail
      Contact( #s60_StWtL1S2DownOver )
      Coil( #qL1S2Down )
   END_RUNG
   // the same network as SCL:
   #qL1S2Down := #s60_StWtL1S2DownOver;
END_REGION

REGION Network 25: Transition for STATE Num:70 StWtOTSFrmConv
   RUNG wire#powerrail
      Contact( #s70_StWtOTSFrmConv )
      I_Contact( #sStWtResetRel )
      Contact( #sSst )
      Contact( #iOTSFrmConv )
      Coil( #s70_StWtOTSFrmConv_T1 )
   END_RUNG
   // the same network as SCL:
   #s70_StWtOTSFrmConv_T1 := #s70_StWtOTSFrmConv AND NOT #sStWtResetRel AND #sSst AND #iOTSFrmConv;
END_REGION

REGION Network 26: STATE Num:70 StWtOTSFrmConv
   RUNG wire#powerrail
      Contact( #s70_StWtOTSFrmConv )
      wire#w1
      I_Contact( #sStWtResetRel )
      I_Contact( #s70_StWtOTSFrmConv_T1 )
      wire#w2
      Coil( #s70_StWtOTSFrmConv )
   END_RUNG
   RUNG wire#powerrail
      Contact( #s60_StWtL1S2DownOver_T1 )
   END_RUNG wire#w1
   RUNG wire#w2
      { S7_GenerateENO := "TRUE" } Move(in := 70, out1 => #StateNo)
   END_RUNG
   // the same network as SCL:
   #s70_StWtOTSFrmConv := (#s70_StWtOTSFrmConv OR #s60_StWtL1S2DownOver_T1) AND NOT #sStWtResetRel AND NOT #s70_StWtOTSFrmConv_T1;
   IF #s70_StWtOTSFrmConv THEN #StateNo := 70; END_IF;
END_REGION

REGION Network 27: Actions for STATE Num:70 StWtOTSFrmConv
   RUNG wire#powerrail
      Contact( #s70_StWtOTSFrmConv )
      Coil( #qRTRToConv )
   END_RUNG
   // the same network as SCL:
   #qRTRToConv := #s70_StWtOTSFrmConv;
END_REGION

REGION Network 28: Transition for STATE Num:80 StWtL1RecvBegin
   RUNG wire#powerrail
      Contact( #s80_StWtL1RecvBegin )
      I_Contact( #sStWtResetRel )
      Contact( #sSst )
      I_Contact( #iAreaClearConv )
      Coil( #s80_StWtL1RecvBegin_T1 )
   END_RUNG
   // the same network as SCL:
   #s80_StWtL1RecvBegin_T1 := #s80_StWtL1RecvBegin AND NOT #sStWtResetRel AND #sSst AND NOT #iAreaClearConv;
END_REGION

REGION Network 29: STATE Num:80 StWtL1RecvBegin
   RUNG wire#powerrail
      Contact( #s80_StWtL1RecvBegin )
      wire#w1
      I_Contact( #sStWtResetRel )
      I_Contact( #s80_StWtL1RecvBegin_T1 )
      wire#w2
      Coil( #s80_StWtL1RecvBegin )
   END_RUNG
   RUNG wire#powerrail
      Contact( #s70_StWtOTSFrmConv_T1 )
   END_RUNG wire#w1
   RUNG wire#w2
      { S7_GenerateENO := "TRUE" } Move(in := 80, out1 => #StateNo)
   END_RUNG
   // the same network as SCL:
   #s80_StWtL1RecvBegin := (#s80_StWtL1RecvBegin OR #s70_StWtOTSFrmConv_T1) AND NOT #sStWtResetRel AND NOT #s80_StWtL1RecvBegin_T1;
   IF #s80_StWtL1RecvBegin THEN #StateNo := 80; END_IF;
END_REGION

REGION Network 30: Transition for STATE Num:90 StWtL1PalRcvDone
   RUNG wire#powerrail
      Contact( #s90_StWtL1PalRcvDone )
      I_Contact( #sStWtResetRel )
      Contact( #sSst )
      Contact( #iL2PalletPrsent )
      Contact( #iAreaClearConv )
      Coil( #s90_StWtL1PalRcvDone_T1 )
   END_RUNG
   // the same network as SCL:
   #s90_StWtL1PalRcvDone_T1 := #s90_StWtL1PalRcvDone AND NOT #sStWtResetRel AND #sSst AND #iL2PalletPrsent AND #iAreaClearConv;
END_REGION

REGION Network 31: STATE Num:90 StWtL1PalRcvDone
   RUNG wire#powerrail
      Contact( #s90_StWtL1PalRcvDone )
      wire#w1
      I_Contact( #sStWtResetRel )
      I_Contact( #s90_StWtL1PalRcvDone_T1 )
      wire#w2
      Coil( #s90_StWtL1PalRcvDone )
   END_RUNG
   RUNG wire#powerrail
      Contact( #s80_StWtL1RecvBegin_T1 )
   END_RUNG wire#w1
   RUNG wire#w2
      { S7_GenerateENO := "TRUE" } Move(in := 90, out1 => #StateNo)
   END_RUNG
   // the same network as SCL:
   #s90_StWtL1PalRcvDone := (#s90_StWtL1PalRcvDone OR #s80_StWtL1RecvBegin_T1) AND NOT #sStWtResetRel AND NOT #s90_StWtL1PalRcvDone_T1;
   IF #s90_StWtL1PalRcvDone THEN #StateNo := 90; END_IF;
END_REGION

REGION Network 32: Transition for STATE Num:100 StRunOutActive
   RUNG wire#powerrail
      Contact( #s100_StRunOutActive )
      I_Contact( #sStWtResetRel )
      Contact( #sSst )
      wire#w1
      I_Contact( #iRunOutCycle )
      Coil( #s100_StRunOutActive_T1 )
   END_RUNG
   RUNG wire#w1
      I_Contact( #s100_StRunOutActive_T1 )
      Contact( #iRunOutCycle )
      Coil( #s100_StRunOutActive_T2 )
   END_RUNG
   // the same network as SCL:
   #_w1 := #s100_StRunOutActive AND NOT #sStWtResetRel AND #sSst;
   #s100_StRunOutActive_T1 := #_w1 AND NOT #iRunOutCycle;
   #s100_StRunOutActive_T2 := #_w1 AND NOT #s100_StRunOutActive_T1 AND #iRunOutCycle;
END_REGION

REGION Network 33: STATE Num:100 StRunOutActive
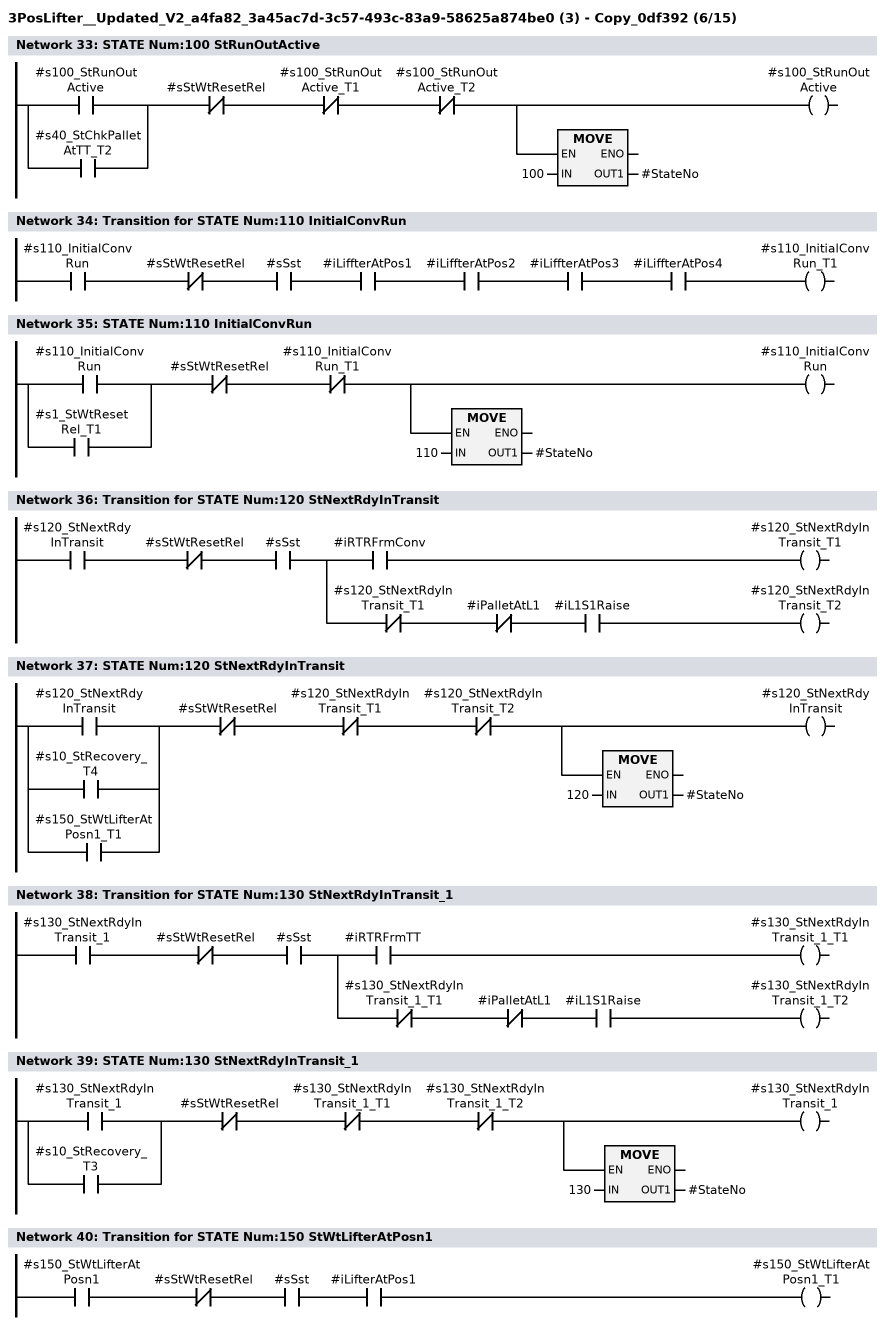
   RUNG wire#powerrail
      Contact( #s100_StRunOutActive )
      wire#w1
      I_Contact( #sStWtResetRel )
      I_Contact( #s100_StRunOutActive_T1 )
      I_Contact( #s100_StRunOutActive_T2 )
      wire#w2
      Coil( #s100_StRunOutActive )
   END_RUNG
   RUNG wire#powerrail
      Contact( #s40_StChkPalletAtTT_T2 )
   END_RUNG wire#w1
   RUNG wire#w2
      { S7_GenerateENO := "TRUE" } Move(in := 100, out1 => #StateNo)
   END_RUNG
   // the same network as SCL:
   #s100_StRunOutActive := (#s100_StRunOutActive OR #s40_StChkPalletAtTT_T2) AND NOT #sStWtResetRel AND NOT #s100_StRunOutActive_T1 AND NOT #s100_StRunOutActive_T2;
   IF #s100_StRunOutActive THEN #StateNo := 100; END_IF;
END_REGION

REGION Network 34: Transition for STATE Num:110 InitialConvRun
   RUNG wire#powerrail
      Contact( #s110_InitialConvRun )
      I_Contact( #sStWtResetRel )
      Contact( #sSst )
      Contact( #iLiffterAtPos1 )
      Contact( #iLiffterAtPos2 )
      Contact( #iLiffterAtPos3 )
      Contact( #iLiffterAtPos4 )
      Coil( #s110_InitialConvRun_T1 )
   END_RUNG
   // the same network as SCL:
   #s110_InitialConvRun_T1 := #s110_InitialConvRun AND NOT #sStWtResetRel AND #sSst AND #iLiffterAtPos1 AND #iLiffterAtPos2 AND #iLiffterAtPos3 AND #iLiffterAtPos4;
END_REGION

REGION Network 35: STATE Num:110 InitialConvRun
   RUNG wire#powerrail
      Contact( #s110_InitialConvRun )
      wire#w1
      I_Contact( #sStWtResetRel )
      I_Contact( #s110_InitialConvRun_T1 )
      wire#w2
      Coil( #s110_InitialConvRun )
   END_RUNG
   RUNG wire#powerrail
      Contact( #s1_StWtResetRel_T1 )
   END_RUNG wire#w1
   RUNG wire#w2
      { S7_GenerateENO := "TRUE" } Move(in := 110, out1 => #StateNo)
   END_RUNG
   // the same network as SCL:
   #s110_InitialConvRun := (#s110_InitialConvRun OR #s1_StWtResetRel_T1) AND NOT #sStWtResetRel AND NOT #s110_InitialConvRun_T1;
   IF #s110_InitialConvRun THEN #StateNo := 110; END_IF;
END_REGION

REGION Network 36: Transition for STATE Num:120 StNextRdyInTransit
   RUNG wire#powerrail
      Contact( #s120_StNextRdyInTransit )
      I_Contact( #sStWtResetRel )
      Contact( #sSst )
      wire#w1
      Contact( #iRTRFrmConv )
      Coil( #s120_StNextRdyInTransit_T1 )
   END_RUNG
   RUNG wire#w1
      I_Contact( #s120_StNextRdyInTransit_T1 )
      I_Contact( #iPalletAtL1 )
      Contact( #iL1S1Raise )
      Coil( #s120_StNextRdyInTransit_T2 )
   END_RUNG
   // the same network as SCL:
   #_w1 := #s120_StNextRdyInTransit AND NOT #sStWtResetRel AND #sSst;
   #s120_StNextRdyInTransit_T1 := #_w1 AND #iRTRFrmConv;
   #s120_StNextRdyInTransit_T2 := #_w1 AND NOT #s120_StNextRdyInTransit_T1 AND NOT #iPalletAtL1 AND #iL1S1Raise;
END_REGION

REGION Network 37: STATE Num:120 StNextRdyInTransit
   RUNG wire#powerrail
      Contact( #s120_StNextRdyInTransit )
      wire#w1
      I_Contact( #sStWtResetRel )
      I_Contact( #s120_StNextRdyInTransit_T1 )
      I_Contact( #s120_StNextRdyInTransit_T2 )
      wire#w2
      Coil( #s120_StNextRdyInTransit )
   END_RUNG
   RUNG wire#powerrail
      Contact( #s10_StRecovery_T4 )
   END_RUNG wire#w1
   RUNG wire#powerrail
      Contact( #s150_StWtLifterAtPosn1_T1 )
   END_RUNG wire#w1
   RUNG wire#w2
      { S7_GenerateENO := "TRUE" } Move(in := 120, out1 => #StateNo)
   END_RUNG
   // the same network as SCL:
   #s120_StNextRdyInTransit := (#s120_StNextRdyInTransit OR #s10_StRecovery_T4 OR #s150_StWtLifterAtPosn1_T1) AND NOT #sStWtResetRel AND NOT #s120_StNextRdyInTransit_T1 AND NOT #s120_StNextRdyInTransit_T2;
   IF #s120_StNextRdyInTransit THEN #StateNo := 120; END_IF;
END_REGION

REGION Network 38: Transition for STATE Num:130 StNextRdyInTransit_1
   RUNG wire#powerrail
      Contact( #s130_StNextRdyInTransit_1 )
      I_Contact( #sStWtResetRel )
      Contact( #sSst )
      wire#w1
      Contact( #iRTRFrmTT )
      Coil( #s130_StNextRdyInTransit_1_T1 )
   END_RUNG
   RUNG wire#w1
      I_Contact( #s130_StNextRdyInTransit_1_T1 )
      I_Contact( #iPalletAtL1 )
      Contact( #iL1S1Raise )
      Coil( #s130_StNextRdyInTransit_1_T2 )
   END_RUNG
   // the same network as SCL:
   #_w1 := #s130_StNextRdyInTransit_1 AND NOT #sStWtResetRel AND #sSst;
   #s130_StNextRdyInTransit_1_T1 := #_w1 AND #iRTRFrmTT;
   #s130_StNextRdyInTransit_1_T2 := #_w1 AND NOT #s130_StNextRdyInTransit_1_T1 AND NOT #iPalletAtL1 AND #iL1S1Raise;
END_REGION

REGION Network 39: STATE Num:130 StNextRdyInTransit_1
   RUNG wire#powerrail
      Contact( #s130_StNextRdyInTransit_1 )
      wire#w1
      I_Contact( #sStWtResetRel )
      I_Contact( #s130_StNextRdyInTransit_1_T1 )
      I_Contact( #s130_StNextRdyInTransit_1_T2 )
      wire#w2
      Coil( #s130_StNextRdyInTransit_1 )
   END_RUNG
   RUNG wire#powerrail
      Contact( #s10_StRecovery_T3 )
   END_RUNG wire#w1
   RUNG wire#w2
      { S7_GenerateENO := "TRUE" } Move(in := 130, out1 => #StateNo)
   END_RUNG
   // the same network as SCL:
   #s130_StNextRdyInTransit_1 := (#s130_StNextRdyInTransit_1 OR #s10_StRecovery_T3) AND NOT #sStWtResetRel AND NOT #s130_StNextRdyInTransit_1_T1 AND NOT #s130_StNextRdyInTransit_1_T2;
   IF #s130_StNextRdyInTransit_1 THEN #StateNo := 130; END_IF;
END_REGION

REGION Network 40: Transition for STATE Num:150 StWtLifterAtPosn1
   RUNG wire#powerrail
      Contact( #s150_StWtLifterAtPosn1 )
      I_Contact( #sStWtResetRel )
      Contact( #sSst )
      Contact( #iLifterAtPos1 )
      Coil( #s150_StWtLifterAtPosn1_T1 )
   END_RUNG
   // the same network as SCL:
   #s150_StWtLifterAtPosn1_T1 := #s150_StWtLifterAtPosn1 AND NOT #sStWtResetRel AND #sSst AND #iLifterAtPos1;
END_REGION

REGION Network 41: STATE Num:150 StWtLifterAtPosn1
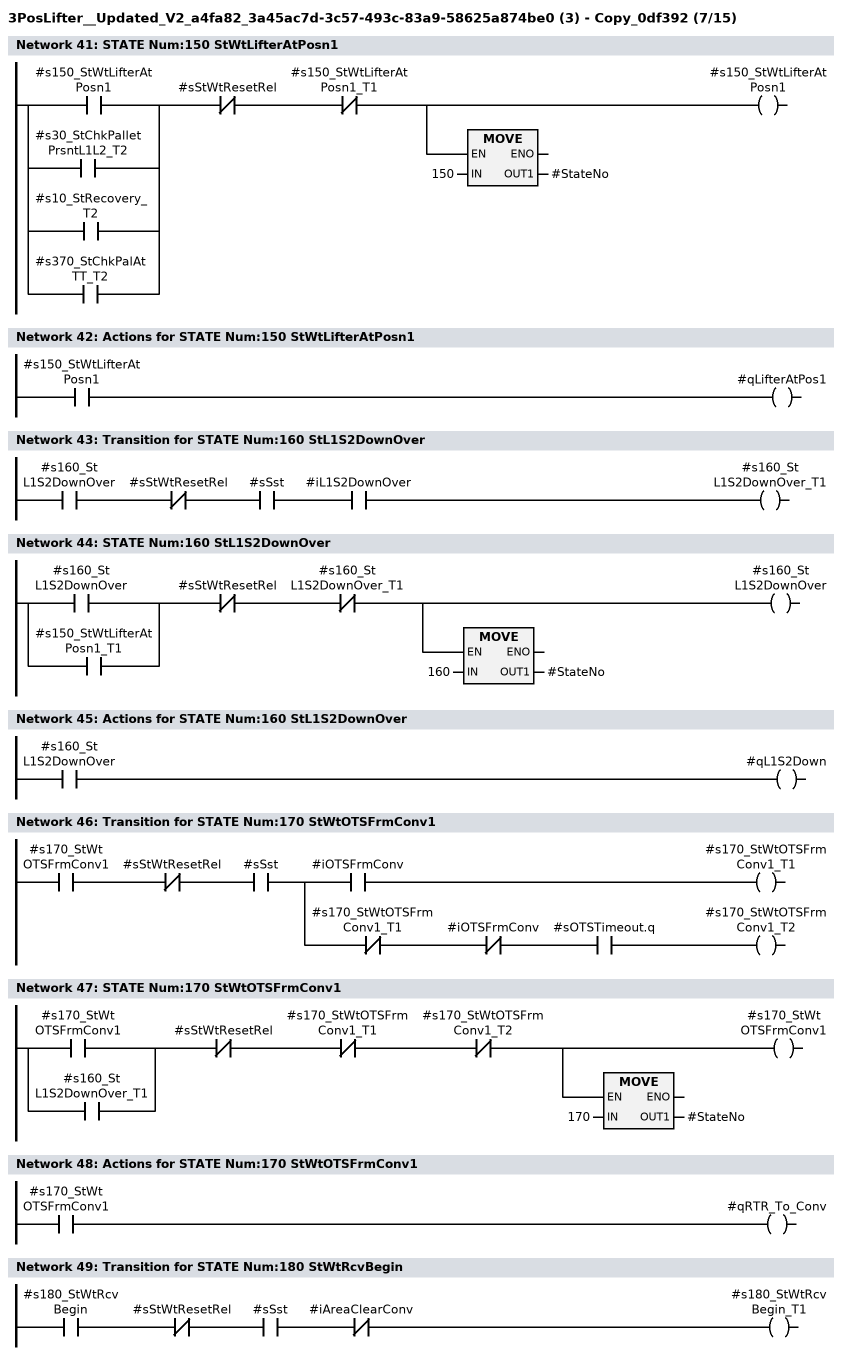
   RUNG wire#powerrail
      Contact( #s150_StWtLifterAtPosn1 )
      wire#w1
      I_Contact( #sStWtResetRel )
      I_Contact( #s150_StWtLifterAtPosn1_T1 )
      wire#w2
      Coil( #s150_StWtLifterAtPosn1 )
   END_RUNG
   RUNG wire#powerrail
      Contact( #s30_StChkPalletPrsntL1L2_T2 )
   END_RUNG wire#w1
   RUNG wire#powerrail
      Contact( #s10_StRecovery_T2 )
   END_RUNG wire#w1
   RUNG wire#powerrail
      Contact( #s370_StChkPalAtTT_T2 )
   END_RUNG wire#w1
   RUNG wire#w2
      { S7_GenerateENO := "TRUE" } Move(in := 150, out1 => #StateNo)
   END_RUNG
   // the same network as SCL:
   #s150_StWtLifterAtPosn1 := (#s150_StWtLifterAtPosn1 OR #s30_StChkPalletPrsntL1L2_T2 OR #s10_StRecovery_T2 OR #s370_StChkPalAtTT_T2) AND NOT #sStWtResetRel AND NOT #s150_StWtLifterAtPosn1_T1;
   IF #s150_StWtLifterAtPosn1 THEN #StateNo := 150; END_IF;
END_REGION

REGION Network 42: Actions for STATE Num:150 StWtLifterAtPosn1
   RUNG wire#powerrail
      Contact( #s150_StWtLifterAtPosn1 )
      Coil( #qLifterAtPos1 )
   END_RUNG
   // the same network as SCL:
   #qLifterAtPos1 := #s150_StWtLifterAtPosn1;
END_REGION

REGION Network 43: Transition for STATE Num:160 StL1S2DownOver
   RUNG wire#powerrail
      Contact( #s160_StL1S2DownOver )
      I_Contact( #sStWtResetRel )
      Contact( #sSst )
      Contact( #iL1S2DownOver )
      Coil( #s160_StL1S2DownOver_T1 )
   END_RUNG
   // the same network as SCL:
   #s160_StL1S2DownOver_T1 := #s160_StL1S2DownOver AND NOT #sStWtResetRel AND #sSst AND #iL1S2DownOver;
END_REGION

REGION Network 44: STATE Num:160 StL1S2DownOver
   RUNG wire#powerrail
      Contact( #s160_StL1S2DownOver )
      wire#w1
      I_Contact( #sStWtResetRel )
      I_Contact( #s160_StL1S2DownOver_T1 )
      wire#w2
      Coil( #s160_StL1S2DownOver )
   END_RUNG
   RUNG wire#powerrail
      Contact( #s150_StWtLifterAtPosn1_T1 )
   END_RUNG wire#w1
   RUNG wire#w2
      { S7_GenerateENO := "TRUE" } Move(in := 160, out1 => #StateNo)
   END_RUNG
   // the same network as SCL:
   #s160_StL1S2DownOver := (#s160_StL1S2DownOver OR #s150_StWtLifterAtPosn1_T1) AND NOT #sStWtResetRel AND NOT #s160_StL1S2DownOver_T1;
   IF #s160_StL1S2DownOver THEN #StateNo := 160; END_IF;
END_REGION

REGION Network 45: Actions for STATE Num:160 StL1S2DownOver
   RUNG wire#powerrail
      Contact( #s160_StL1S2DownOver )
      Coil( #qL1S2Down )
   END_RUNG
   // the same network as SCL:
   #qL1S2Down := #s160_StL1S2DownOver;
END_REGION

REGION Network 46: Transition for STATE Num:170 StWtOTSFrmConv1
   RUNG wire#powerrail
      Contact( #s170_StWtOTSFrmConv1 )
      I_Contact( #sStWtResetRel )
      Contact( #sSst )
      wire#w1
      Contact( #iOTSFrmConv )
      Coil( #s170_StWtOTSFrmConv1_T1 )
   END_RUNG
   RUNG wire#w1
      I_Contact( #s170_StWtOTSFrmConv1_T1 )
      I_Contact( #iOTSFrmConv )
      Contact( #sOTSTimeout.q )
      Coil( #s170_StWtOTSFrmConv1_T2 )
   END_RUNG
   // the same network as SCL:
   #_w1 := #s170_StWtOTSFrmConv1 AND NOT #sStWtResetRel AND #sSst;
   #s170_StWtOTSFrmConv1_T1 := #_w1 AND #iOTSFrmConv;
   #s170_StWtOTSFrmConv1_T2 := #_w1 AND NOT #s170_StWtOTSFrmConv1_T1 AND NOT #iOTSFrmConv AND #sOTSTimeout.q;
END_REGION

REGION Network 47: STATE Num:170 StWtOTSFrmConv1
   RUNG wire#powerrail
      Contact( #s170_StWtOTSFrmConv1 )
      wire#w1
      I_Contact( #sStWtResetRel )
      I_Contact( #s170_StWtOTSFrmConv1_T1 )
      I_Contact( #s170_StWtOTSFrmConv1_T2 )
      wire#w2
      Coil( #s170_StWtOTSFrmConv1 )
   END_RUNG
   RUNG wire#powerrail
      Contact( #s160_StL1S2DownOver_T1 )
   END_RUNG wire#w1
   RUNG wire#w2
      { S7_GenerateENO := "TRUE" } Move(in := 170, out1 => #StateNo)
   END_RUNG
   // the same network as SCL:
   #s170_StWtOTSFrmConv1 := (#s170_StWtOTSFrmConv1 OR #s160_StL1S2DownOver_T1) AND NOT #sStWtResetRel AND NOT #s170_StWtOTSFrmConv1_T1 AND NOT #s170_StWtOTSFrmConv1_T2;
   IF #s170_StWtOTSFrmConv1 THEN #StateNo := 170; END_IF;
END_REGION

REGION Network 48: Actions for STATE Num:170 StWtOTSFrmConv1
   RUNG wire#powerrail
      Contact( #s170_StWtOTSFrmConv1 )
      Coil( #qRTR_To_Conv )
   END_RUNG
   // the same network as SCL:
   #qRTR_To_Conv := #s170_StWtOTSFrmConv1;
END_REGION

REGION Network 49: Transition for STATE Num:180 StWtRcvBegin
   RUNG wire#powerrail
      Contact( #s180_StWtRcvBegin )
      I_Contact( #sStWtResetRel )
      Contact( #sSst )
      I_Contact( #iAreaClearConv )
      Coil( #s180_StWtRcvBegin_T1 )
   END_RUNG
   // the same network as SCL:
   #s180_StWtRcvBegin_T1 := #s180_StWtRcvBegin AND NOT #sStWtResetRel AND #sSst AND NOT #iAreaClearConv;
END_REGION

REGION Network 50: STATE Num:180 StWtRcvBegin
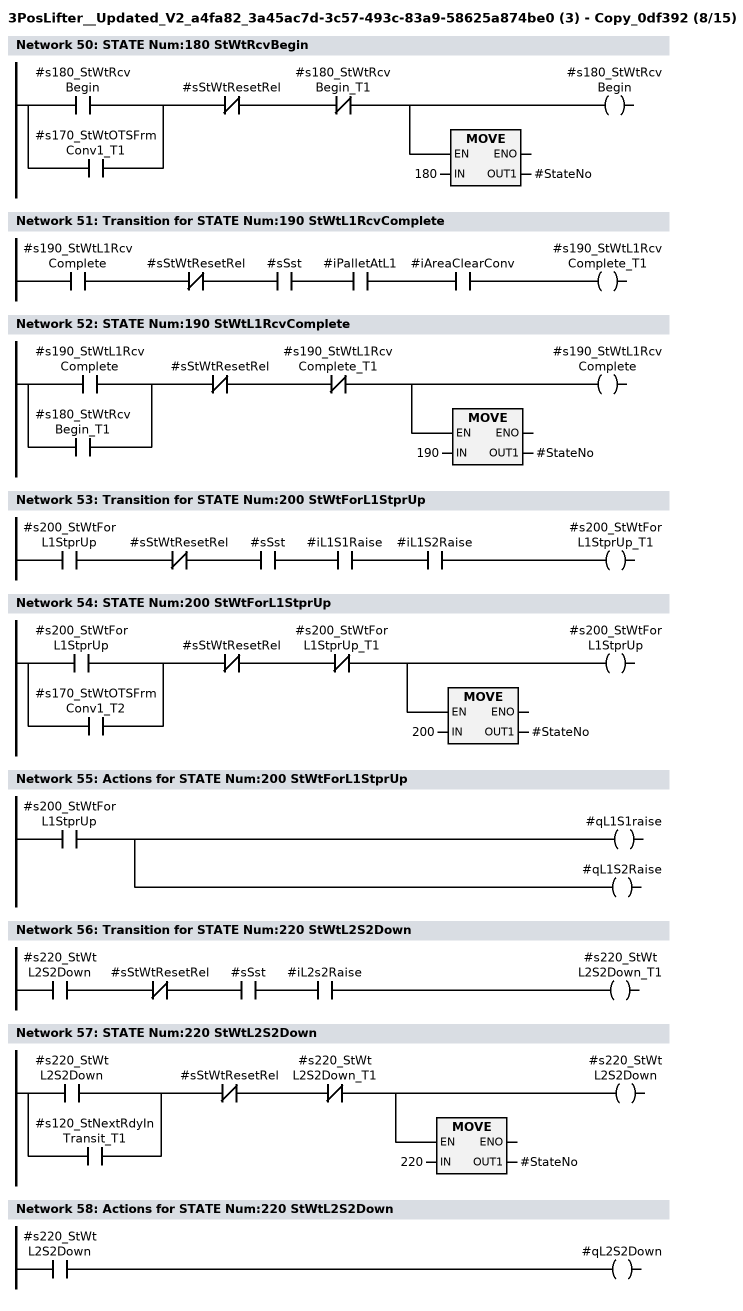
   RUNG wire#powerrail
      Contact( #s180_StWtRcvBegin )
      wire#w1
      I_Contact( #sStWtResetRel )
      I_Contact( #s180_StWtRcvBegin_T1 )
      wire#w2
      Coil( #s180_StWtRcvBegin )
   END_RUNG
   RUNG wire#powerrail
      Contact( #s170_StWtOTSFrmConv1_T1 )
   END_RUNG wire#w1
   RUNG wire#w2
      { S7_GenerateENO := "TRUE" } Move(in := 180, out1 => #StateNo)
   END_RUNG
   // the same network as SCL:
   #s180_StWtRcvBegin := (#s180_StWtRcvBegin OR #s170_StWtOTSFrmConv1_T1) AND NOT #sStWtResetRel AND NOT #s180_StWtRcvBegin_T1;
   IF #s180_StWtRcvBegin THEN #StateNo := 180; END_IF;
END_REGION

REGION Network 51: Transition for STATE Num:190 StWtL1RcvComplete
   RUNG wire#powerrail
      Contact( #s190_StWtL1RcvComplete )
      I_Contact( #sStWtResetRel )
      Contact( #sSst )
      Contact( #iPalletAtL1 )
      Contact( #iAreaClearConv )
      Coil( #s190_StWtL1RcvComplete_T1 )
   END_RUNG
   // the same network as SCL:
   #s190_StWtL1RcvComplete_T1 := #s190_StWtL1RcvComplete AND NOT #sStWtResetRel AND #sSst AND #iPalletAtL1 AND #iAreaClearConv;
END_REGION

REGION Network 52: STATE Num:190 StWtL1RcvComplete
   RUNG wire#powerrail
      Contact( #s190_StWtL1RcvComplete )
      wire#w1
      I_Contact( #sStWtResetRel )
      I_Contact( #s190_StWtL1RcvComplete_T1 )
      wire#w2
      Coil( #s190_StWtL1RcvComplete )
   END_RUNG
   RUNG wire#powerrail
      Contact( #s180_StWtRcvBegin_T1 )
   END_RUNG wire#w1
   RUNG wire#w2
      { S7_GenerateENO := "TRUE" } Move(in := 190, out1 => #StateNo)
   END_RUNG
   // the same network as SCL:
   #s190_StWtL1RcvComplete := (#s190_StWtL1RcvComplete OR #s180_StWtRcvBegin_T1) AND NOT #sStWtResetRel AND NOT #s190_StWtL1RcvComplete_T1;
   IF #s190_StWtL1RcvComplete THEN #StateNo := 190; END_IF;
END_REGION

REGION Network 53: Transition for STATE Num:200 StWtForL1StprUp
   RUNG wire#powerrail
      Contact( #s200_StWtForL1StprUp )
      I_Contact( #sStWtResetRel )
      Contact( #sSst )
      Contact( #iL1S1Raise )
      Contact( #iL1S2Raise )
      Coil( #s200_StWtForL1StprUp_T1 )
   END_RUNG
   // the same network as SCL:
   #s200_StWtForL1StprUp_T1 := #s200_StWtForL1StprUp AND NOT #sStWtResetRel AND #sSst AND #iL1S1Raise AND #iL1S2Raise;
END_REGION

REGION Network 54: STATE Num:200 StWtForL1StprUp
   RUNG wire#powerrail
      Contact( #s200_StWtForL1StprUp )
      wire#w1
      I_Contact( #sStWtResetRel )
      I_Contact( #s200_StWtForL1StprUp_T1 )
      wire#w2
      Coil( #s200_StWtForL1StprUp )
   END_RUNG
   RUNG wire#powerrail
      Contact( #s170_StWtOTSFrmConv1_T2 )
   END_RUNG wire#w1
   RUNG wire#w2
      { S7_GenerateENO := "TRUE" } Move(in := 200, out1 => #StateNo)
   END_RUNG
   // the same network as SCL:
   #s200_StWtForL1StprUp := (#s200_StWtForL1StprUp OR #s170_StWtOTSFrmConv1_T2) AND NOT #sStWtResetRel AND NOT #s200_StWtForL1StprUp_T1;
   IF #s200_StWtForL1StprUp THEN #StateNo := 200; END_IF;
END_REGION

REGION Network 55: Actions for STATE Num:200 StWtForL1StprUp
   RUNG wire#powerrail
      Contact( #s200_StWtForL1StprUp )
      wire#w1
      Coil( #qL1S1raise )
   END_RUNG
   RUNG wire#w1
      Coil( #qL1S2Raise )
   END_RUNG
   // the same network as SCL:
   #qL1S1raise := #s200_StWtForL1StprUp;
   #qL1S2Raise := #s200_StWtForL1StprUp;
END_REGION

REGION Network 56: Transition for STATE Num:220 StWtL2S2Down
   RUNG wire#powerrail
      Contact( #s220_StWtL2S2Down )
      I_Contact( #sStWtResetRel )
      Contact( #sSst )
      Contact( #iL2s2Raise )
      Coil( #s220_StWtL2S2Down_T1 )
   END_RUNG
   // the same network as SCL:
   #s220_StWtL2S2Down_T1 := #s220_StWtL2S2Down AND NOT #sStWtResetRel AND #sSst AND #iL2s2Raise;
END_REGION

REGION Network 57: STATE Num:220 StWtL2S2Down
   RUNG wire#powerrail
      Contact( #s220_StWtL2S2Down )
      wire#w1
      I_Contact( #sStWtResetRel )
      I_Contact( #s220_StWtL2S2Down_T1 )
      wire#w2
      Coil( #s220_StWtL2S2Down )
   END_RUNG
   RUNG wire#powerrail
      Contact( #s120_StNextRdyInTransit_T1 )
   END_RUNG wire#w1
   RUNG wire#w2
      { S7_GenerateENO := "TRUE" } Move(in := 220, out1 => #StateNo)
   END_RUNG
   // the same network as SCL:
   #s220_StWtL2S2Down := (#s220_StWtL2S2Down OR #s120_StNextRdyInTransit_T1) AND NOT #sStWtResetRel AND NOT #s220_StWtL2S2Down_T1;
   IF #s220_StWtL2S2Down THEN #StateNo := 220; END_IF;
END_REGION

REGION Network 58: Actions for STATE Num:220 StWtL2S2Down
   RUNG wire#powerrail
      Contact( #s220_StWtL2S2Down )
      Coil( #qL2S2Down )
   END_RUNG
   // the same network as SCL:
   #qL2S2Down := #s220_StWtL2S2Down;
END_REGION

REGION Network 59: Transition for STATE Num:230 StWtL2TranBegin
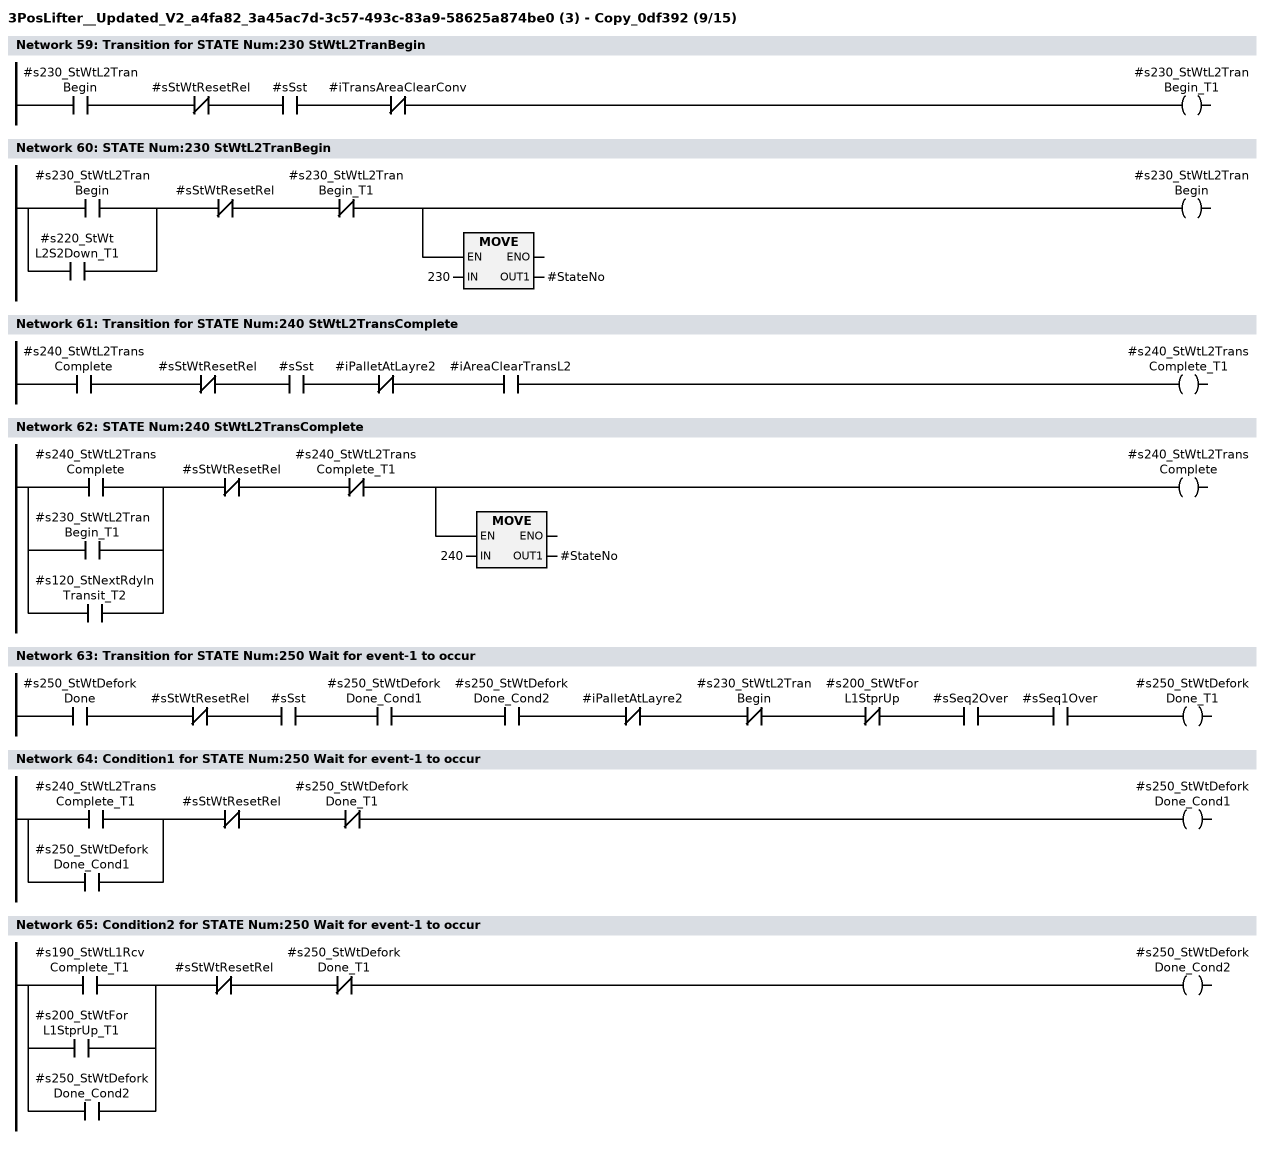
   RUNG wire#powerrail
      Contact( #s230_StWtL2TranBegin )
      I_Contact( #sStWtResetRel )
      Contact( #sSst )
      I_Contact( #iTransAreaClearConv )
      Coil( #s230_StWtL2TranBegin_T1 )
   END_RUNG
   // the same network as SCL:
   #s230_StWtL2TranBegin_T1 := #s230_StWtL2TranBegin AND NOT #sStWtResetRel AND #sSst AND NOT #iTransAreaClearConv;
END_REGION

REGION Network 60: STATE Num:230 StWtL2TranBegin
   RUNG wire#powerrail
      Contact( #s230_StWtL2TranBegin )
      wire#w1
      I_Contact( #sStWtResetRel )
      I_Contact( #s230_StWtL2TranBegin_T1 )
      wire#w2
      Coil( #s230_StWtL2TranBegin )
   END_RUNG
   RUNG wire#powerrail
      Contact( #s220_StWtL2S2Down_T1 )
   END_RUNG wire#w1
   RUNG wire#w2
      { S7_GenerateENO := "TRUE" } Move(in := 230, out1 => #StateNo)
   END_RUNG
   // the same network as SCL:
   #s230_StWtL2TranBegin := (#s230_StWtL2TranBegin OR #s220_StWtL2S2Down_T1) AND NOT #sStWtResetRel AND NOT #s230_StWtL2TranBegin_T1;
   IF #s230_StWtL2TranBegin THEN #StateNo := 230; END_IF;
END_REGION

REGION Network 61: Transition for STATE Num:240 StWtL2TransComplete
   RUNG wire#powerrail
      Contact( #s240_StWtL2TransComplete )
      I_Contact( #sStWtResetRel )
      Contact( #sSst )
      I_Contact( #iPalletAtLayre2 )
      Contact( #iAreaClearTransL2 )
      Coil( #s240_StWtL2TransComplete_T1 )
   END_RUNG
   // the same network as SCL:
   #s240_StWtL2TransComplete_T1 := #s240_StWtL2TransComplete AND NOT #sStWtResetRel AND #sSst AND NOT #iPalletAtLayre2 AND #iAreaClearTransL2;
END_REGION

REGION Network 62: STATE Num:240 StWtL2TransComplete
   RUNG wire#powerrail
      Contact( #s240_StWtL2TransComplete )
      wire#w1
      I_Contact( #sStWtResetRel )
      I_Contact( #s240_StWtL2TransComplete_T1 )
      wire#w2
      Coil( #s240_StWtL2TransComplete )
   END_RUNG
   RUNG wire#powerrail
      Contact( #s230_StWtL2TranBegin_T1 )
   END_RUNG wire#w1
   RUNG wire#powerrail
      Contact( #s120_StNextRdyInTransit_T2 )
   END_RUNG wire#w1
   RUNG wire#w2
      { S7_GenerateENO := "TRUE" } Move(in := 240, out1 => #StateNo)
   END_RUNG
   // the same network as SCL:
   #s240_StWtL2TransComplete := (#s240_StWtL2TransComplete OR #s230_StWtL2TranBegin_T1 OR #s120_StNextRdyInTransit_T2) AND NOT #sStWtResetRel AND NOT #s240_StWtL2TransComplete_T1;
   IF #s240_StWtL2TransComplete THEN #StateNo := 240; END_IF;
END_REGION

REGION Network 63: Transition for STATE Num:250 Wait for event-1 to occur
   RUNG wire#powerrail
      Contact( #s250_StWtDeforkDone )
      I_Contact( #sStWtResetRel )
      Contact( #sSst )
      Contact( #s250_StWtDeforkDone_Cond1 )
      Contact( #s250_StWtDeforkDone_Cond2 )
      I_Contact( #iPalletAtLayre2 )
      I_Contact( #s230_StWtL2TranBegin )
      I_Contact( #s200_StWtForL1StprUp )
      Contact( #sSeq2Over )
      Contact( #sSeq1Over )
      Coil( #s250_StWtDeforkDone_T1 )
   END_RUNG
   // the same network as SCL:
   #s250_StWtDeforkDone_T1 := #s250_StWtDeforkDone AND NOT #sStWtResetRel AND #sSst AND #s250_StWtDeforkDone_Cond1 AND #s250_StWtDeforkDone_Cond2 AND NOT #iPalletAtLayre2 AND NOT #s230_StWtL2TranBegin AND NOT #s200_StWtForL1StprUp AND #sSeq2Over AND #sSeq1Over;
END_REGION

REGION Network 64: Condition1 for STATE Num:250 Wait for event-1 to occur
   RUNG wire#powerrail
      Contact( #s240_StWtL2TransComplete_T1 )
      wire#w1
      I_Contact( #sStWtResetRel )
      I_Contact( #s250_StWtDeforkDone_T1 )
      Coil( #s250_StWtDeforkDone_Cond1 )
   END_RUNG
   RUNG wire#powerrail
      Contact( #s250_StWtDeforkDone_Cond1 )
   END_RUNG wire#w1
   // the same network as SCL:
   #s250_StWtDeforkDone_Cond1 := (#s240_StWtL2TransComplete_T1 OR #s250_StWtDeforkDone_Cond1) AND NOT #sStWtResetRel AND NOT #s250_StWtDeforkDone_T1;
END_REGION

REGION Network 65: Condition2 for STATE Num:250 Wait for event-1 to occur
   RUNG wire#powerrail
      Contact( #s190_StWtL1RcvComplete_T1 )
      wire#w1
      I_Contact( #sStWtResetRel )
      I_Contact( #s250_StWtDeforkDone_T1 )
      Coil( #s250_StWtDeforkDone_Cond2 )
   END_RUNG
   RUNG wire#powerrail
      Contact( #s200_StWtForL1StprUp_T1 )
   END_RUNG wire#w1
   RUNG wire#powerrail
      Contact( #s250_StWtDeforkDone_Cond2 )
   END_RUNG wire#w1
   // the same network as SCL:
   #s250_StWtDeforkDone_Cond2 := (#s190_StWtL1RcvComplete_T1 OR #s200_StWtForL1StprUp_T1 OR #s250_StWtDeforkDone_Cond2) AND NOT #sStWtResetRel AND NOT #s250_StWtDeforkDone_T1;
END_REGION

REGION Network 66: STATE Num:250 Wait for event-1 to occur
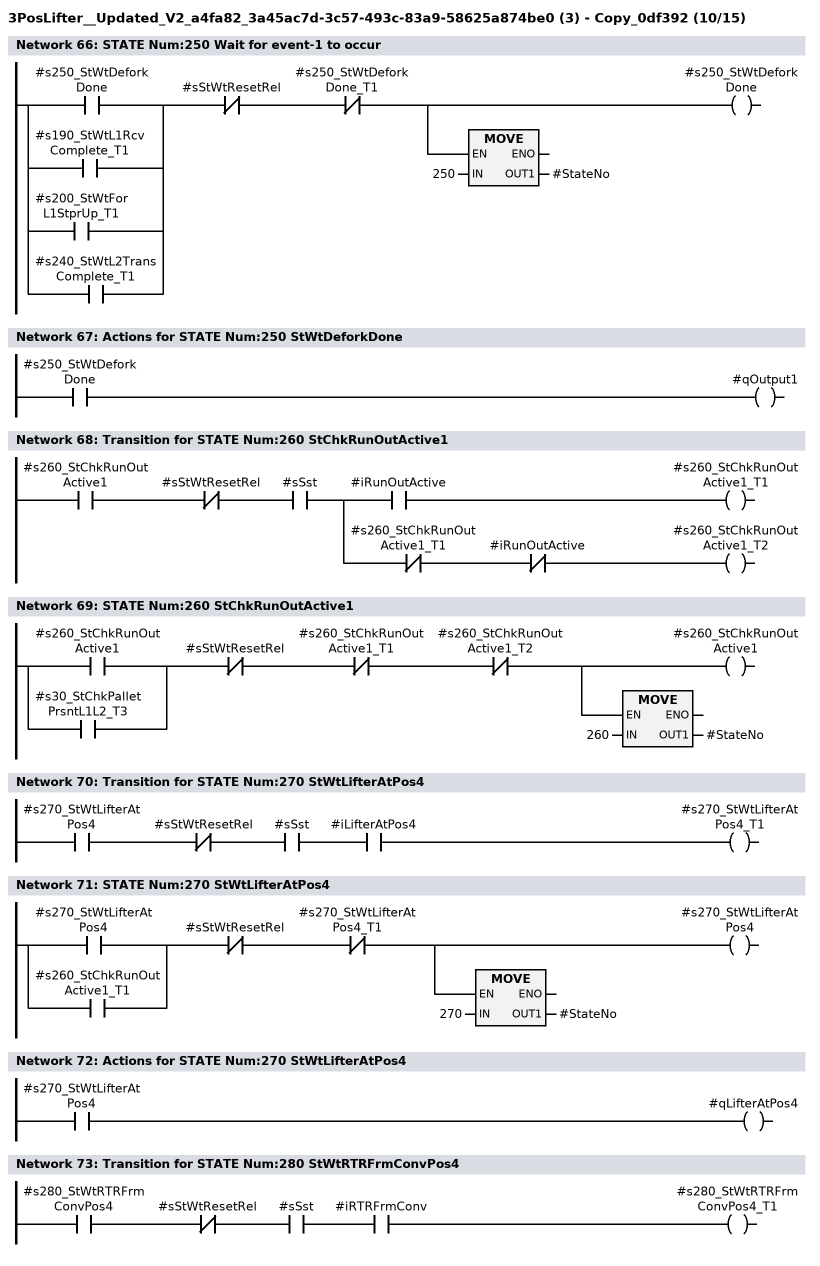
   RUNG wire#powerrail
      Contact( #s250_StWtDeforkDone )
      wire#w1
      I_Contact( #sStWtResetRel )
      I_Contact( #s250_StWtDeforkDone_T1 )
      wire#w2
      Coil( #s250_StWtDeforkDone )
   END_RUNG
   RUNG wire#powerrail
      Contact( #s190_StWtL1RcvComplete_T1 )
   END_RUNG wire#w1
   RUNG wire#powerrail
      Contact( #s200_StWtForL1StprUp_T1 )
   END_RUNG wire#w1
   RUNG wire#powerrail
      Contact( #s240_StWtL2TransComplete_T1 )
   END_RUNG wire#w1
   RUNG wire#w2
      { S7_GenerateENO := "TRUE" } Move(in := 250, out1 => #StateNo)
   END_RUNG
   // the same network as SCL:
   #s250_StWtDeforkDone := (#s250_StWtDeforkDone OR #s190_StWtL1RcvComplete_T1 OR #s200_StWtForL1StprUp_T1 OR #s240_StWtL2TransComplete_T1) AND NOT #sStWtResetRel AND NOT #s250_StWtDeforkDone_T1;
   IF #s250_StWtDeforkDone THEN #StateNo := 250; END_IF;
END_REGION

REGION Network 67: Actions for STATE Num:250 StWtDeforkDone
   RUNG wire#powerrail
      Contact( #s250_StWtDeforkDone )
      Coil( #qOutput1 )
   END_RUNG
   // the same network as SCL:
   #qOutput1 := #s250_StWtDeforkDone;
END_REGION

REGION Network 68: Transition for STATE Num:260 StChkRunOutActive1
   RUNG wire#powerrail
      Contact( #s260_StChkRunOutActive1 )
      I_Contact( #sStWtResetRel )
      Contact( #sSst )
      wire#w1
      Contact( #iRunOutActive )
      Coil( #s260_StChkRunOutActive1_T1 )
   END_RUNG
   RUNG wire#w1
      I_Contact( #s260_StChkRunOutActive1_T1 )
      I_Contact( #iRunOutActive )
      Coil( #s260_StChkRunOutActive1_T2 )
   END_RUNG
   // the same network as SCL:
   #_w1 := #s260_StChkRunOutActive1 AND NOT #sStWtResetRel AND #sSst;
   #s260_StChkRunOutActive1_T1 := #_w1 AND #iRunOutActive;
   #s260_StChkRunOutActive1_T2 := #_w1 AND NOT #s260_StChkRunOutActive1_T1 AND NOT #iRunOutActive;
END_REGION

REGION Network 69: STATE Num:260 StChkRunOutActive1
   RUNG wire#powerrail
      Contact( #s260_StChkRunOutActive1 )
      wire#w1
      I_Contact( #sStWtResetRel )
      I_Contact( #s260_StChkRunOutActive1_T1 )
      I_Contact( #s260_StChkRunOutActive1_T2 )
      wire#w2
      Coil( #s260_StChkRunOutActive1 )
   END_RUNG
   RUNG wire#powerrail
      Contact( #s30_StChkPalletPrsntL1L2_T3 )
   END_RUNG wire#w1
   RUNG wire#w2
      { S7_GenerateENO := "TRUE" } Move(in := 260, out1 => #StateNo)
   END_RUNG
   // the same network as SCL:
   #s260_StChkRunOutActive1 := (#s260_StChkRunOutActive1 OR #s30_StChkPalletPrsntL1L2_T3) AND NOT #sStWtResetRel AND NOT #s260_StChkRunOutActive1_T1 AND NOT #s260_StChkRunOutActive1_T2;
   IF #s260_StChkRunOutActive1 THEN #StateNo := 260; END_IF;
END_REGION

REGION Network 70: Transition for STATE Num:270 StWtLifterAtPos4
   RUNG wire#powerrail
      Contact( #s270_StWtLifterAtPos4 )
      I_Contact( #sStWtResetRel )
      Contact( #sSst )
      Contact( #iLifterAtPos4 )
      Coil( #s270_StWtLifterAtPos4_T1 )
   END_RUNG
   // the same network as SCL:
   #s270_StWtLifterAtPos4_T1 := #s270_StWtLifterAtPos4 AND NOT #sStWtResetRel AND #sSst AND #iLifterAtPos4;
END_REGION

REGION Network 71: STATE Num:270 StWtLifterAtPos4
   RUNG wire#powerrail
      Contact( #s270_StWtLifterAtPos4 )
      wire#w1
      I_Contact( #sStWtResetRel )
      I_Contact( #s270_StWtLifterAtPos4_T1 )
      wire#w2
      Coil( #s270_StWtLifterAtPos4 )
   END_RUNG
   RUNG wire#powerrail
      Contact( #s260_StChkRunOutActive1_T1 )
   END_RUNG wire#w1
   RUNG wire#w2
      { S7_GenerateENO := "TRUE" } Move(in := 270, out1 => #StateNo)
   END_RUNG
   // the same network as SCL:
   #s270_StWtLifterAtPos4 := (#s270_StWtLifterAtPos4 OR #s260_StChkRunOutActive1_T1) AND NOT #sStWtResetRel AND NOT #s270_StWtLifterAtPos4_T1;
   IF #s270_StWtLifterAtPos4 THEN #StateNo := 270; END_IF;
END_REGION

REGION Network 72: Actions for STATE Num:270 StWtLifterAtPos4
   RUNG wire#powerrail
      Contact( #s270_StWtLifterAtPos4 )
      Coil( #qLifterAtPos4 )
   END_RUNG
   // the same network as SCL:
   #qLifterAtPos4 := #s270_StWtLifterAtPos4;
END_REGION

REGION Network 73: Transition for STATE Num:280 StWtRTRFrmConvPos4
   RUNG wire#powerrail
      Contact( #s280_StWtRTRFrmConvPos4 )
      I_Contact( #sStWtResetRel )
      Contact( #sSst )
      Contact( #iRTRFrmConv )
      Coil( #s280_StWtRTRFrmConvPos4_T1 )
   END_RUNG
   // the same network as SCL:
   #s280_StWtRTRFrmConvPos4_T1 := #s280_StWtRTRFrmConvPos4 AND NOT #sStWtResetRel AND #sSst AND #iRTRFrmConv;
END_REGION

REGION Network 74: STATE Num:280 StWtRTRFrmConvPos4
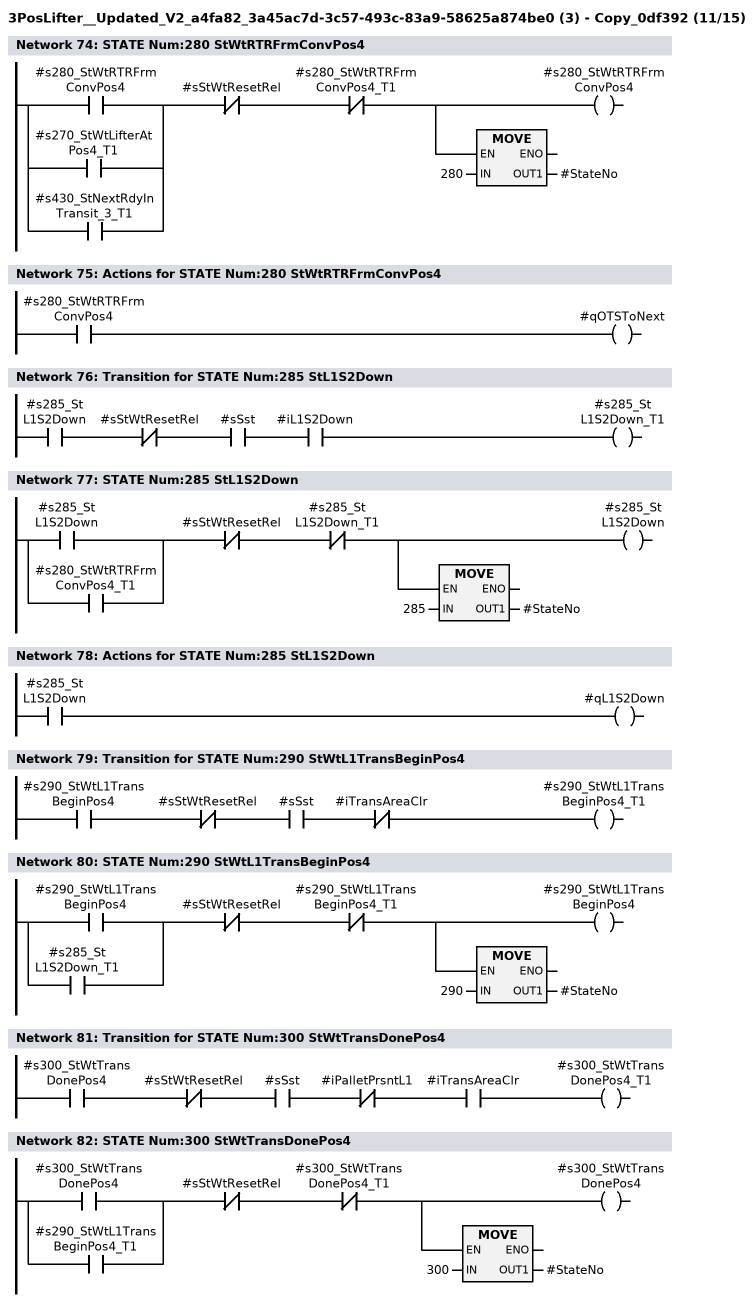
   RUNG wire#powerrail
      Contact( #s280_StWtRTRFrmConvPos4 )
      wire#w1
      I_Contact( #sStWtResetRel )
      I_Contact( #s280_StWtRTRFrmConvPos4_T1 )
      wire#w2
      Coil( #s280_StWtRTRFrmConvPos4 )
   END_RUNG
   RUNG wire#powerrail
      Contact( #s270_StWtLifterAtPos4_T1 )
   END_RUNG wire#w1
   RUNG wire#powerrail
      Contact( #s430_StNextRdyInTransit_3_T1 )
   END_RUNG wire#w1
   RUNG wire#w2
      { S7_GenerateENO := "TRUE" } Move(in := 280, out1 => #StateNo)
   END_RUNG
   // the same network as SCL:
   #s280_StWtRTRFrmConvPos4 := (#s280_StWtRTRFrmConvPos4 OR #s270_StWtLifterAtPos4_T1 OR #s430_StNextRdyInTransit_3_T1) AND NOT #sStWtResetRel AND NOT #s280_StWtRTRFrmConvPos4_T1;
   IF #s280_StWtRTRFrmConvPos4 THEN #StateNo := 280; END_IF;
END_REGION

REGION Network 75: Actions for STATE Num:280 StWtRTRFrmConvPos4
   RUNG wire#powerrail
      Contact( #s280_StWtRTRFrmConvPos4 )
      Coil( #qOTSToNext )
   END_RUNG
   // the same network as SCL:
   #qOTSToNext := #s280_StWtRTRFrmConvPos4;
END_REGION

REGION Network 76: Transition for STATE Num:285 StL1S2Down
   RUNG wire#powerrail
      Contact( #s285_StL1S2Down )
      I_Contact( #sStWtResetRel )
      Contact( #sSst )
      Contact( #iL1S2Down )
      Coil( #s285_StL1S2Down_T1 )
   END_RUNG
   // the same network as SCL:
   #s285_StL1S2Down_T1 := #s285_StL1S2Down AND NOT #sStWtResetRel AND #sSst AND #iL1S2Down;
END_REGION

REGION Network 77: STATE Num:285 StL1S2Down
   RUNG wire#powerrail
      Contact( #s285_StL1S2Down )
      wire#w1
      I_Contact( #sStWtResetRel )
      I_Contact( #s285_StL1S2Down_T1 )
      wire#w2
      Coil( #s285_StL1S2Down )
   END_RUNG
   RUNG wire#powerrail
      Contact( #s280_StWtRTRFrmConvPos4_T1 )
   END_RUNG wire#w1
   RUNG wire#w2
      { S7_GenerateENO := "TRUE" } Move(in := 285, out1 => #StateNo)
   END_RUNG
   // the same network as SCL:
   #s285_StL1S2Down := (#s285_StL1S2Down OR #s280_StWtRTRFrmConvPos4_T1) AND NOT #sStWtResetRel AND NOT #s285_StL1S2Down_T1;
   IF #s285_StL1S2Down THEN #StateNo := 285; END_IF;
END_REGION

REGION Network 78: Actions for STATE Num:285 StL1S2Down
   RUNG wire#powerrail
      Contact( #s285_StL1S2Down )
      Coil( #qL1S2Down )
   END_RUNG
   // the same network as SCL:
   #qL1S2Down := #s285_StL1S2Down;
END_REGION

REGION Network 79: Transition for STATE Num:290 StWtL1TransBeginPos4
   RUNG wire#powerrail
      Contact( #s290_StWtL1TransBeginPos4 )
      I_Contact( #sStWtResetRel )
      Contact( #sSst )
      I_Contact( #iTransAreaClr )
      Coil( #s290_StWtL1TransBeginPos4_T1 )
   END_RUNG
   // the same network as SCL:
   #s290_StWtL1TransBeginPos4_T1 := #s290_StWtL1TransBeginPos4 AND NOT #sStWtResetRel AND #sSst AND NOT #iTransAreaClr;
END_REGION

REGION Network 80: STATE Num:290 StWtL1TransBeginPos4
   RUNG wire#powerrail
      Contact( #s290_StWtL1TransBeginPos4 )
      wire#w1
      I_Contact( #sStWtResetRel )
      I_Contact( #s290_StWtL1TransBeginPos4_T1 )
      wire#w2
      Coil( #s290_StWtL1TransBeginPos4 )
   END_RUNG
   RUNG wire#powerrail
      Contact( #s285_StL1S2Down_T1 )
   END_RUNG wire#w1
   RUNG wire#w2
      { S7_GenerateENO := "TRUE" } Move(in := 290, out1 => #StateNo)
   END_RUNG
   // the same network as SCL:
   #s290_StWtL1TransBeginPos4 := (#s290_StWtL1TransBeginPos4 OR #s285_StL1S2Down_T1) AND NOT #sStWtResetRel AND NOT #s290_StWtL1TransBeginPos4_T1;
   IF #s290_StWtL1TransBeginPos4 THEN #StateNo := 290; END_IF;
END_REGION

REGION Network 81: Transition for STATE Num:300 StWtTransDonePos4
   RUNG wire#powerrail
      Contact( #s300_StWtTransDonePos4 )
      I_Contact( #sStWtResetRel )
      Contact( #sSst )
      I_Contact( #iPalletPrsntL1 )
      Contact( #iTransAreaClr )
      Coil( #s300_StWtTransDonePos4_T1 )
   END_RUNG
   // the same network as SCL:
   #s300_StWtTransDonePos4_T1 := #s300_StWtTransDonePos4 AND NOT #sStWtResetRel AND #sSst AND NOT #iPalletPrsntL1 AND #iTransAreaClr;
END_REGION

REGION Network 82: STATE Num:300 StWtTransDonePos4
   RUNG wire#powerrail
      Contact( #s300_StWtTransDonePos4 )
      wire#w1
      I_Contact( #sStWtResetRel )
      I_Contact( #s300_StWtTransDonePos4_T1 )
      wire#w2
      Coil( #s300_StWtTransDonePos4 )
   END_RUNG
   RUNG wire#powerrail
      Contact( #s290_StWtL1TransBeginPos4_T1 )
   END_RUNG wire#w1
   RUNG wire#w2
      { S7_GenerateENO := "TRUE" } Move(in := 300, out1 => #StateNo)
   END_RUNG
   // the same network as SCL:
   #s300_StWtTransDonePos4 := (#s300_StWtTransDonePos4 OR #s290_StWtL1TransBeginPos4_T1) AND NOT #sStWtResetRel AND NOT #s300_StWtTransDonePos4_T1;
   IF #s300_StWtTransDonePos4 THEN #StateNo := 300; END_IF;
END_REGION

REGION Network 83: Transition for STATE Num:310 StChkPalletAtTT1
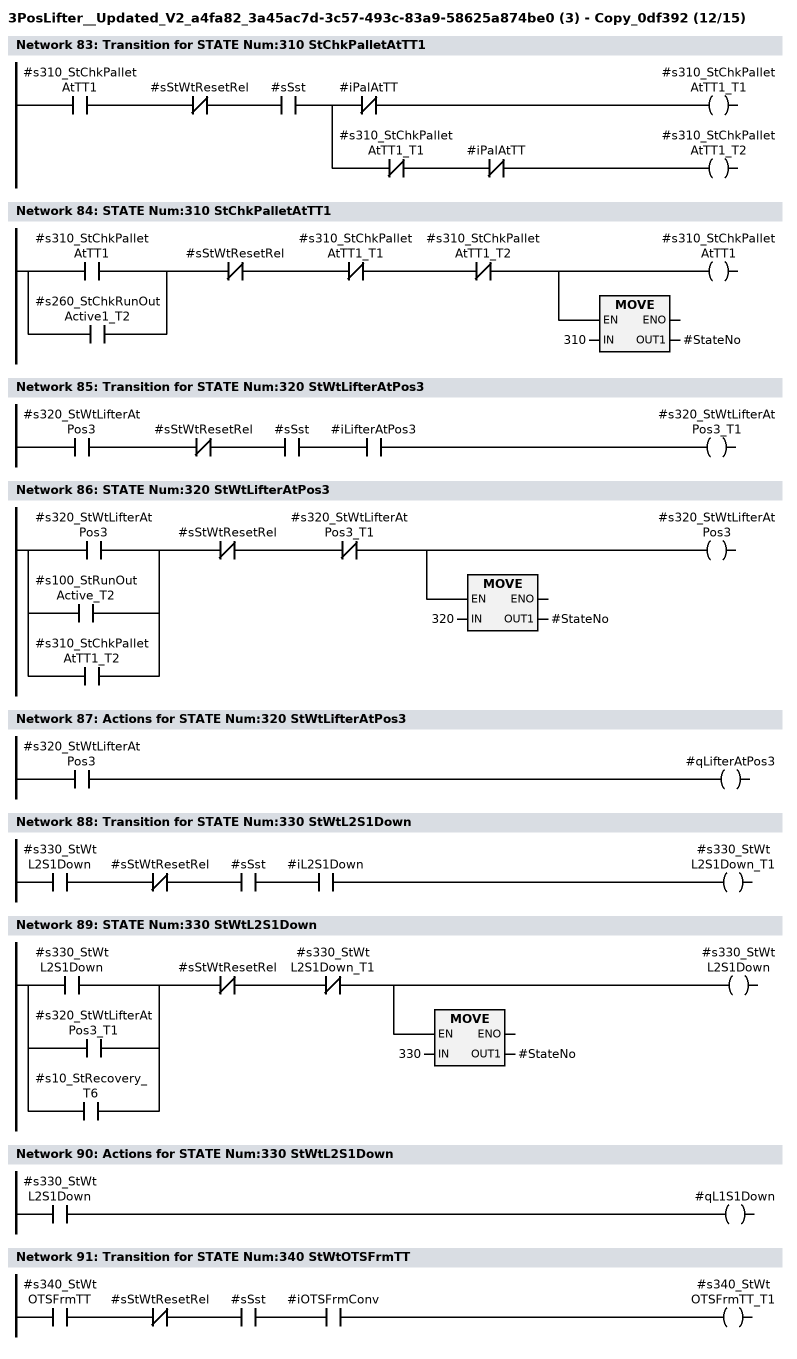
   RUNG wire#powerrail
      Contact( #s310_StChkPalletAtTT1 )
      I_Contact( #sStWtResetRel )
      Contact( #sSst )
      wire#w1
      I_Contact( #iPalAtTT )
      Coil( #s310_StChkPalletAtTT1_T1 )
   END_RUNG
   RUNG wire#w1
      I_Contact( #s310_StChkPalletAtTT1_T1 )
      I_Contact( #iPalAtTT )
      Coil( #s310_StChkPalletAtTT1_T2 )
   END_RUNG
   // the same network as SCL:
   #_w1 := #s310_StChkPalletAtTT1 AND NOT #sStWtResetRel AND #sSst;
   #s310_StChkPalletAtTT1_T1 := #_w1 AND NOT #iPalAtTT;
   #s310_StChkPalletAtTT1_T2 := #_w1 AND NOT #s310_StChkPalletAtTT1_T1 AND NOT #iPalAtTT;
END_REGION

REGION Network 84: STATE Num:310 StChkPalletAtTT1
   RUNG wire#powerrail
      Contact( #s310_StChkPalletAtTT1 )
      wire#w1
      I_Contact( #sStWtResetRel )
      I_Contact( #s310_StChkPalletAtTT1_T1 )
      I_Contact( #s310_StChkPalletAtTT1_T2 )
      wire#w2
      Coil( #s310_StChkPalletAtTT1 )
   END_RUNG
   RUNG wire#powerrail
      Contact( #s260_StChkRunOutActive1_T2 )
   END_RUNG wire#w1
   RUNG wire#w2
      { S7_GenerateENO := "TRUE" } Move(in := 310, out1 => #StateNo)
   END_RUNG
   // the same network as SCL:
   #s310_StChkPalletAtTT1 := (#s310_StChkPalletAtTT1 OR #s260_StChkRunOutActive1_T2) AND NOT #sStWtResetRel AND NOT #s310_StChkPalletAtTT1_T1 AND NOT #s310_StChkPalletAtTT1_T2;
   IF #s310_StChkPalletAtTT1 THEN #StateNo := 310; END_IF;
END_REGION

REGION Network 85: Transition for STATE Num:320 StWtLifterAtPos3
   RUNG wire#powerrail
      Contact( #s320_StWtLifterAtPos3 )
      I_Contact( #sStWtResetRel )
      Contact( #sSst )
      Contact( #iLifterAtPos3 )
      Coil( #s320_StWtLifterAtPos3_T1 )
   END_RUNG
   // the same network as SCL:
   #s320_StWtLifterAtPos3_T1 := #s320_StWtLifterAtPos3 AND NOT #sStWtResetRel AND #sSst AND #iLifterAtPos3;
END_REGION

REGION Network 86: STATE Num:320 StWtLifterAtPos3
   RUNG wire#powerrail
      Contact( #s320_StWtLifterAtPos3 )
      wire#w1
      I_Contact( #sStWtResetRel )
      I_Contact( #s320_StWtLifterAtPos3_T1 )
      wire#w2
      Coil( #s320_StWtLifterAtPos3 )
   END_RUNG
   RUNG wire#powerrail
      Contact( #s100_StRunOutActive_T2 )
   END_RUNG wire#w1
   RUNG wire#powerrail
      Contact( #s310_StChkPalletAtTT1_T2 )
   END_RUNG wire#w1
   RUNG wire#w2
      { S7_GenerateENO := "TRUE" } Move(in := 320, out1 => #StateNo)
   END_RUNG
   // the same network as SCL:
   #s320_StWtLifterAtPos3 := (#s320_StWtLifterAtPos3 OR #s100_StRunOutActive_T2 OR #s310_StChkPalletAtTT1_T2) AND NOT #sStWtResetRel AND NOT #s320_StWtLifterAtPos3_T1;
   IF #s320_StWtLifterAtPos3 THEN #StateNo := 320; END_IF;
END_REGION

REGION Network 87: Actions for STATE Num:320 StWtLifterAtPos3
   RUNG wire#powerrail
      Contact( #s320_StWtLifterAtPos3 )
      Coil( #qLifterAtPos3 )
   END_RUNG
   // the same network as SCL:
   #qLifterAtPos3 := #s320_StWtLifterAtPos3;
END_REGION

REGION Network 88: Transition for STATE Num:330 StWtL2S1Down
   RUNG wire#powerrail
      Contact( #s330_StWtL2S1Down )
      I_Contact( #sStWtResetRel )
      Contact( #sSst )
      Contact( #iL2S1Down )
      Coil( #s330_StWtL2S1Down_T1 )
   END_RUNG
   // the same network as SCL:
   #s330_StWtL2S1Down_T1 := #s330_StWtL2S1Down AND NOT #sStWtResetRel AND #sSst AND #iL2S1Down;
END_REGION

REGION Network 89: STATE Num:330 StWtL2S1Down
   RUNG wire#powerrail
      Contact( #s330_StWtL2S1Down )
      wire#w1
      I_Contact( #sStWtResetRel )
      I_Contact( #s330_StWtL2S1Down_T1 )
      wire#w2
      Coil( #s330_StWtL2S1Down )
   END_RUNG
   RUNG wire#powerrail
      Contact( #s320_StWtLifterAtPos3_T1 )
   END_RUNG wire#w1
   RUNG wire#powerrail
      Contact( #s10_StRecovery_T6 )
   END_RUNG wire#w1
   RUNG wire#w2
      { S7_GenerateENO := "TRUE" } Move(in := 330, out1 => #StateNo)
   END_RUNG
   // the same network as SCL:
   #s330_StWtL2S1Down := (#s330_StWtL2S1Down OR #s320_StWtLifterAtPos3_T1 OR #s10_StRecovery_T6) AND NOT #sStWtResetRel AND NOT #s330_StWtL2S1Down_T1;
   IF #s330_StWtL2S1Down THEN #StateNo := 330; END_IF;
END_REGION

REGION Network 90: Actions for STATE Num:330 StWtL2S1Down
   RUNG wire#powerrail
      Contact( #s330_StWtL2S1Down )
      Coil( #qL1S1Down )
   END_RUNG
   // the same network as SCL:
   #qL1S1Down := #s330_StWtL2S1Down;
END_REGION

REGION Network 91: Transition for STATE Num:340 StWtOTSFrmTT
   RUNG wire#powerrail
      Contact( #s340_StWtOTSFrmTT )
      I_Contact( #sStWtResetRel )
      Contact( #sSst )
      Contact( #iOTSFrmConv )
      Coil( #s340_StWtOTSFrmTT_T1 )
   END_RUNG
   // the same network as SCL:
   #s340_StWtOTSFrmTT_T1 := #s340_StWtOTSFrmTT AND NOT #sStWtResetRel AND #sSst AND #iOTSFrmConv;
END_REGION

REGION Network 92: STATE Num:340 StWtOTSFrmTT
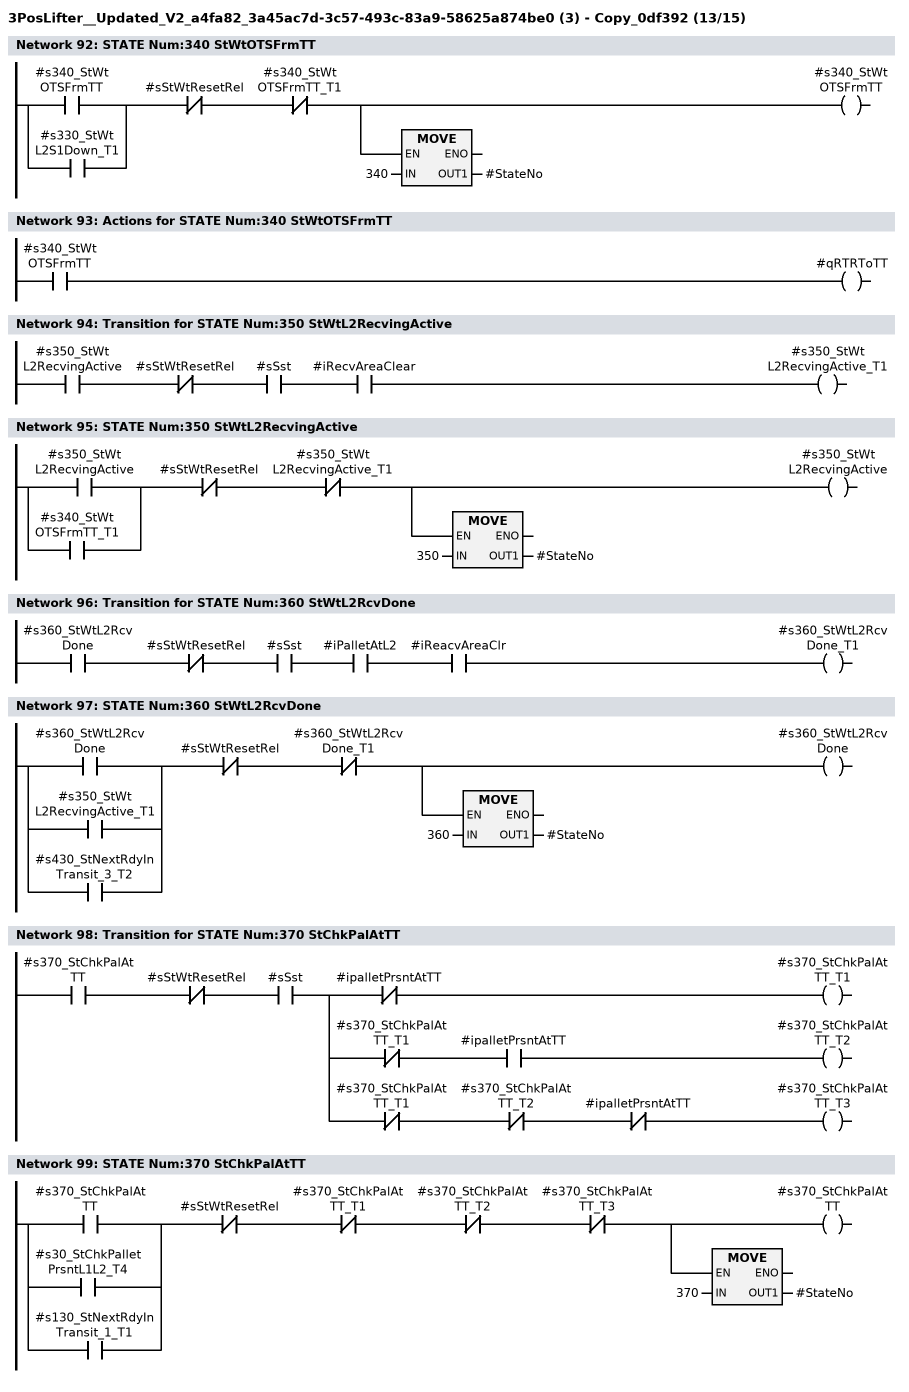
   RUNG wire#powerrail
      Contact( #s340_StWtOTSFrmTT )
      wire#w1
      I_Contact( #sStWtResetRel )
      I_Contact( #s340_StWtOTSFrmTT_T1 )
      wire#w2
      Coil( #s340_StWtOTSFrmTT )
   END_RUNG
   RUNG wire#powerrail
      Contact( #s330_StWtL2S1Down_T1 )
   END_RUNG wire#w1
   RUNG wire#w2
      { S7_GenerateENO := "TRUE" } Move(in := 340, out1 => #StateNo)
   END_RUNG
   // the same network as SCL:
   #s340_StWtOTSFrmTT := (#s340_StWtOTSFrmTT OR #s330_StWtL2S1Down_T1) AND NOT #sStWtResetRel AND NOT #s340_StWtOTSFrmTT_T1;
   IF #s340_StWtOTSFrmTT THEN #StateNo := 340; END_IF;
END_REGION

REGION Network 93: Actions for STATE Num:340 StWtOTSFrmTT
   RUNG wire#powerrail
      Contact( #s340_StWtOTSFrmTT )
      Coil( #qRTRToTT )
   END_RUNG
   // the same network as SCL:
   #qRTRToTT := #s340_StWtOTSFrmTT;
END_REGION

REGION Network 94: Transition for STATE Num:350 StWtL2RecvingActive
   RUNG wire#powerrail
      Contact( #s350_StWtL2RecvingActive )
      I_Contact( #sStWtResetRel )
      Contact( #sSst )
      Contact( #iRecvAreaClear )
      Coil( #s350_StWtL2RecvingActive_T1 )
   END_RUNG
   // the same network as SCL:
   #s350_StWtL2RecvingActive_T1 := #s350_StWtL2RecvingActive AND NOT #sStWtResetRel AND #sSst AND #iRecvAreaClear;
END_REGION

REGION Network 95: STATE Num:350 StWtL2RecvingActive
   RUNG wire#powerrail
      Contact( #s350_StWtL2RecvingActive )
      wire#w1
      I_Contact( #sStWtResetRel )
      I_Contact( #s350_StWtL2RecvingActive_T1 )
      wire#w2
      Coil( #s350_StWtL2RecvingActive )
   END_RUNG
   RUNG wire#powerrail
      Contact( #s340_StWtOTSFrmTT_T1 )
   END_RUNG wire#w1
   RUNG wire#w2
      { S7_GenerateENO := "TRUE" } Move(in := 350, out1 => #StateNo)
   END_RUNG
   // the same network as SCL:
   #s350_StWtL2RecvingActive := (#s350_StWtL2RecvingActive OR #s340_StWtOTSFrmTT_T1) AND NOT #sStWtResetRel AND NOT #s350_StWtL2RecvingActive_T1;
   IF #s350_StWtL2RecvingActive THEN #StateNo := 350; END_IF;
END_REGION

REGION Network 96: Transition for STATE Num:360 StWtL2RcvDone
   RUNG wire#powerrail
      Contact( #s360_StWtL2RcvDone )
      I_Contact( #sStWtResetRel )
      Contact( #sSst )
      Contact( #iPalletAtL2 )
      Contact( #iReacvAreaClr )
      Coil( #s360_StWtL2RcvDone_T1 )
   END_RUNG
   // the same network as SCL:
   #s360_StWtL2RcvDone_T1 := #s360_StWtL2RcvDone AND NOT #sStWtResetRel AND #sSst AND #iPalletAtL2 AND #iReacvAreaClr;
END_REGION

REGION Network 97: STATE Num:360 StWtL2RcvDone
   RUNG wire#powerrail
      Contact( #s360_StWtL2RcvDone )
      wire#w1
      I_Contact( #sStWtResetRel )
      I_Contact( #s360_StWtL2RcvDone_T1 )
      wire#w2
      Coil( #s360_StWtL2RcvDone )
   END_RUNG
   RUNG wire#powerrail
      Contact( #s350_StWtL2RecvingActive_T1 )
   END_RUNG wire#w1
   RUNG wire#powerrail
      Contact( #s430_StNextRdyInTransit_3_T2 )
   END_RUNG wire#w1
   RUNG wire#w2
      { S7_GenerateENO := "TRUE" } Move(in := 360, out1 => #StateNo)
   END_RUNG
   // the same network as SCL:
   #s360_StWtL2RcvDone := (#s360_StWtL2RcvDone OR #s350_StWtL2RecvingActive_T1 OR #s430_StNextRdyInTransit_3_T2) AND NOT #sStWtResetRel AND NOT #s360_StWtL2RcvDone_T1;
   IF #s360_StWtL2RcvDone THEN #StateNo := 360; END_IF;
END_REGION

REGION Network 98: Transition for STATE Num:370 StChkPalAtTT
   RUNG wire#powerrail
      Contact( #s370_StChkPalAtTT )
      I_Contact( #sStWtResetRel )
      Contact( #sSst )
      wire#w1
      I_Contact( #ipalletPrsntAtTT )
      Coil( #s370_StChkPalAtTT_T1 )
   END_RUNG
   RUNG wire#w1
      I_Contact( #s370_StChkPalAtTT_T1 )
      Contact( #ipalletPrsntAtTT )
      Coil( #s370_StChkPalAtTT_T2 )
   END_RUNG
   RUNG wire#w1
      I_Contact( #s370_StChkPalAtTT_T1 )
      I_Contact( #s370_StChkPalAtTT_T2 )
      I_Contact( #ipalletPrsntAtTT )
      Coil( #s370_StChkPalAtTT_T3 )
   END_RUNG
   // the same network as SCL:
   #_w1 := #s370_StChkPalAtTT AND NOT #sStWtResetRel AND #sSst;
   #s370_StChkPalAtTT_T1 := #_w1 AND NOT #ipalletPrsntAtTT;
   #s370_StChkPalAtTT_T2 := #_w1 AND NOT #s370_StChkPalAtTT_T1 AND #ipalletPrsntAtTT;
   #s370_StChkPalAtTT_T3 := #_w1 AND NOT #s370_StChkPalAtTT_T1 AND NOT #s370_StChkPalAtTT_T2 AND NOT #ipalletPrsntAtTT;
END_REGION

REGION Network 99: STATE Num:370 StChkPalAtTT
   RUNG wire#powerrail
      Contact( #s370_StChkPalAtTT )
      wire#w1
      I_Contact( #sStWtResetRel )
      I_Contact( #s370_StChkPalAtTT_T1 )
      I_Contact( #s370_StChkPalAtTT_T2 )
      I_Contact( #s370_StChkPalAtTT_T3 )
      wire#w2
      Coil( #s370_StChkPalAtTT )
   END_RUNG
   RUNG wire#powerrail
      Contact( #s30_StChkPalletPrsntL1L2_T4 )
   END_RUNG wire#w1
   RUNG wire#powerrail
      Contact( #s130_StNextRdyInTransit_1_T1 )
   END_RUNG wire#w1
   RUNG wire#w2
      { S7_GenerateENO := "TRUE" } Move(in := 370, out1 => #StateNo)
   END_RUNG
   // the same network as SCL:
   #s370_StChkPalAtTT := (#s370_StChkPalAtTT OR #s30_StChkPalletPrsntL1L2_T4 OR #s130_StNextRdyInTransit_1_T1) AND NOT #sStWtResetRel AND NOT #s370_StChkPalAtTT_T1 AND NOT #s370_StChkPalAtTT_T2 AND NOT #s370_StChkPalAtTT_T3;
   IF #s370_StChkPalAtTT THEN #StateNo := 370; END_IF;
END_REGION

REGION Network 100: Transition for STATE Num:380 StWtLifterAtPos2
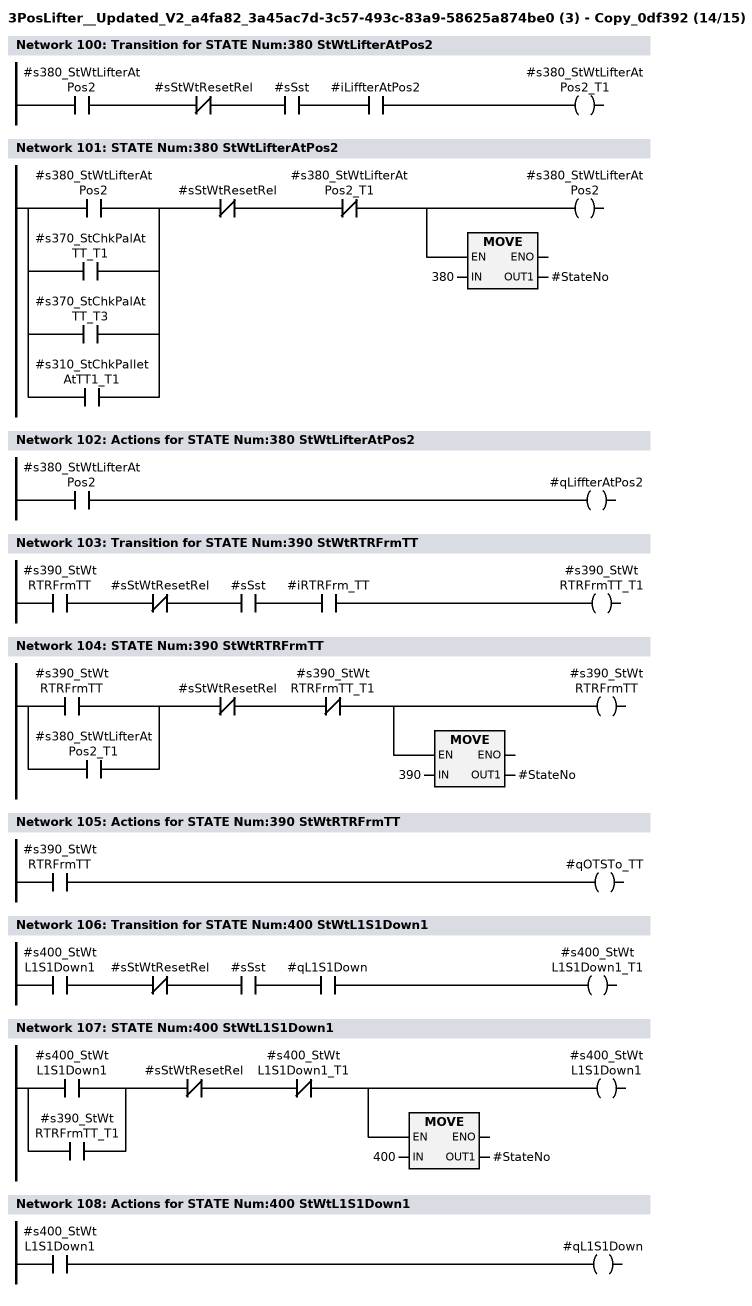
   RUNG wire#powerrail
      Contact( #s380_StWtLifterAtPos2 )
      I_Contact( #sStWtResetRel )
      Contact( #sSst )
      Contact( #iLiffterAtPos2 )
      Coil( #s380_StWtLifterAtPos2_T1 )
   END_RUNG
   // the same network as SCL:
   #s380_StWtLifterAtPos2_T1 := #s380_StWtLifterAtPos2 AND NOT #sStWtResetRel AND #sSst AND #iLiffterAtPos2;
END_REGION

REGION Network 101: STATE Num:380 StWtLifterAtPos2
   RUNG wire#powerrail
      Contact( #s380_StWtLifterAtPos2 )
      wire#w1
      I_Contact( #sStWtResetRel )
      I_Contact( #s380_StWtLifterAtPos2_T1 )
      wire#w2
      Coil( #s380_StWtLifterAtPos2 )
   END_RUNG
   RUNG wire#powerrail
      Contact( #s370_StChkPalAtTT_T1 )
   END_RUNG wire#w1
   RUNG wire#powerrail
      Contact( #s370_StChkPalAtTT_T3 )
   END_RUNG wire#w1
   RUNG wire#powerrail
      Contact( #s310_StChkPalletAtTT1_T1 )
   END_RUNG wire#w1
   RUNG wire#w2
      { S7_GenerateENO := "TRUE" } Move(in := 380, out1 => #StateNo)
   END_RUNG
   // the same network as SCL:
   #s380_StWtLifterAtPos2 := (#s380_StWtLifterAtPos2 OR #s370_StChkPalAtTT_T1 OR #s370_StChkPalAtTT_T3 OR #s310_StChkPalletAtTT1_T1) AND NOT #sStWtResetRel AND NOT #s380_StWtLifterAtPos2_T1;
   IF #s380_StWtLifterAtPos2 THEN #StateNo := 380; END_IF;
END_REGION

REGION Network 102: Actions for STATE Num:380 StWtLifterAtPos2
   RUNG wire#powerrail
      Contact( #s380_StWtLifterAtPos2 )
      Coil( #qLiffterAtPos2 )
   END_RUNG
   // the same network as SCL:
   #qLiffterAtPos2 := #s380_StWtLifterAtPos2;
END_REGION

REGION Network 103: Transition for STATE Num:390 StWtRTRFrmTT
   RUNG wire#powerrail
      Contact( #s390_StWtRTRFrmTT )
      I_Contact( #sStWtResetRel )
      Contact( #sSst )
      Contact( #iRTRFrm_TT )
      Coil( #s390_StWtRTRFrmTT_T1 )
   END_RUNG
   // the same network as SCL:
   #s390_StWtRTRFrmTT_T1 := #s390_StWtRTRFrmTT AND NOT #sStWtResetRel AND #sSst AND #iRTRFrm_TT;
END_REGION

REGION Network 104: STATE Num:390 StWtRTRFrmTT
   RUNG wire#powerrail
      Contact( #s390_StWtRTRFrmTT )
      wire#w1
      I_Contact( #sStWtResetRel )
      I_Contact( #s390_StWtRTRFrmTT_T1 )
      wire#w2
      Coil( #s390_StWtRTRFrmTT )
   END_RUNG
   RUNG wire#powerrail
      Contact( #s380_StWtLifterAtPos2_T1 )
   END_RUNG wire#w1
   RUNG wire#w2
      { S7_GenerateENO := "TRUE" } Move(in := 390, out1 => #StateNo)
   END_RUNG
   // the same network as SCL:
   #s390_StWtRTRFrmTT := (#s390_StWtRTRFrmTT OR #s380_StWtLifterAtPos2_T1) AND NOT #sStWtResetRel AND NOT #s390_StWtRTRFrmTT_T1;
   IF #s390_StWtRTRFrmTT THEN #StateNo := 390; END_IF;
END_REGION

REGION Network 105: Actions for STATE Num:390 StWtRTRFrmTT
   RUNG wire#powerrail
      Contact( #s390_StWtRTRFrmTT )
      Coil( #qOTSTo_TT )
   END_RUNG
   // the same network as SCL:
   #qOTSTo_TT := #s390_StWtRTRFrmTT;
END_REGION

REGION Network 106: Transition for STATE Num:400 StWtL1S1Down1
   RUNG wire#powerrail
      Contact( #s400_StWtL1S1Down1 )
      I_Contact( #sStWtResetRel )
      Contact( #sSst )
      Contact( #qL1S1Down )
      Coil( #s400_StWtL1S1Down1_T1 )
   END_RUNG
   // the same network as SCL:
   #s400_StWtL1S1Down1_T1 := #s400_StWtL1S1Down1 AND NOT #sStWtResetRel AND #sSst AND #qL1S1Down;
END_REGION

REGION Network 107: STATE Num:400 StWtL1S1Down1
   RUNG wire#powerrail
      Contact( #s400_StWtL1S1Down1 )
      wire#w1
      I_Contact( #sStWtResetRel )
      I_Contact( #s400_StWtL1S1Down1_T1 )
      wire#w2
      Coil( #s400_StWtL1S1Down1 )
   END_RUNG
   RUNG wire#powerrail
      Contact( #s390_StWtRTRFrmTT_T1 )
   END_RUNG wire#w1
   RUNG wire#w2
      { S7_GenerateENO := "TRUE" } Move(in := 400, out1 => #StateNo)
   END_RUNG
   // the same network as SCL:
   #s400_StWtL1S1Down1 := (#s400_StWtL1S1Down1 OR #s390_StWtRTRFrmTT_T1) AND NOT #sStWtResetRel AND NOT #s400_StWtL1S1Down1_T1;
   IF #s400_StWtL1S1Down1 THEN #StateNo := 400; END_IF;
END_REGION

REGION Network 108: Actions for STATE Num:400 StWtL1S1Down1
   RUNG wire#powerrail
      Contact( #s400_StWtL1S1Down1 )
      Coil( #qL1S1Down )
   END_RUNG
   // the same network as SCL:
   #qL1S1Down := #s400_StWtL1S1Down1;
END_REGION

REGION Network 109: Transition for STATE Num:410 StWtL1TransBegin
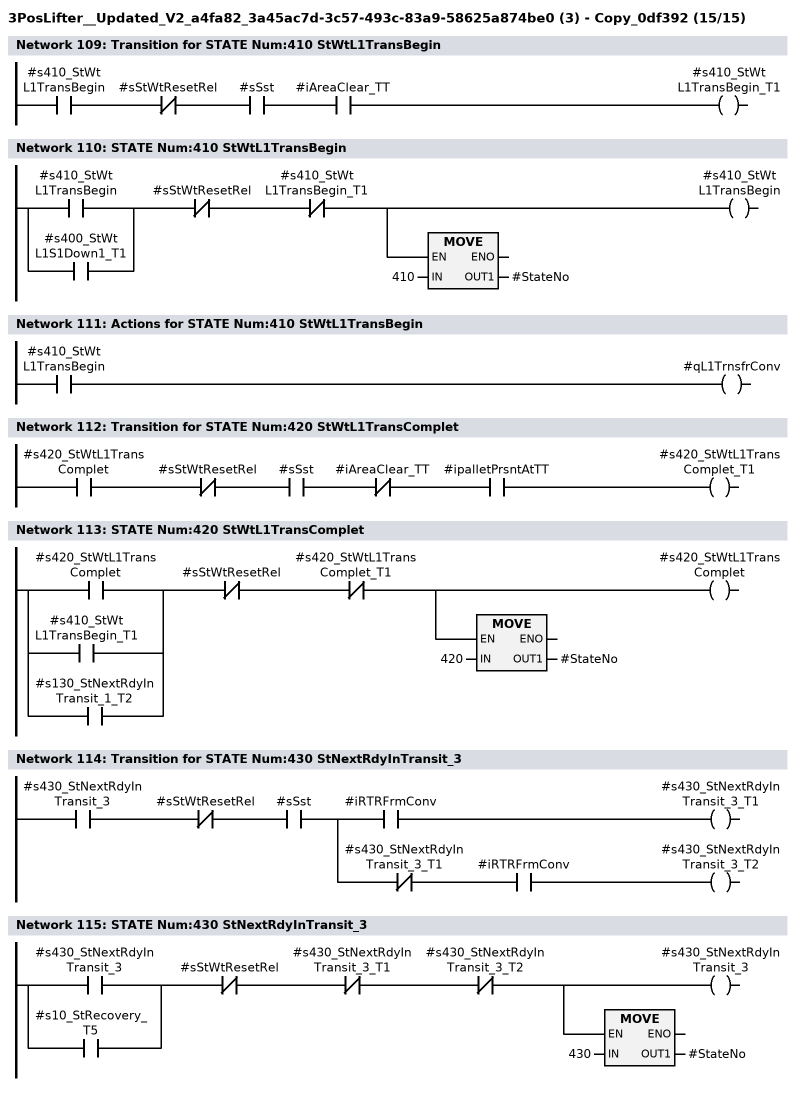
   RUNG wire#powerrail
      Contact( #s410_StWtL1TransBegin )
      I_Contact( #sStWtResetRel )
      Contact( #sSst )
      Contact( #iAreaClear_TT )
      Coil( #s410_StWtL1TransBegin_T1 )
   END_RUNG
   // the same network as SCL:
   #s410_StWtL1TransBegin_T1 := #s410_StWtL1TransBegin AND NOT #sStWtResetRel AND #sSst AND #iAreaClear_TT;
END_REGION

REGION Network 110: STATE Num:410 StWtL1TransBegin
   RUNG wire#powerrail
      Contact( #s410_StWtL1TransBegin )
      wire#w1
      I_Contact( #sStWtResetRel )
      I_Contact( #s410_StWtL1TransBegin_T1 )
      wire#w2
      Coil( #s410_StWtL1TransBegin )
   END_RUNG
   RUNG wire#powerrail
      Contact( #s400_StWtL1S1Down1_T1 )
   END_RUNG wire#w1
   RUNG wire#w2
      { S7_GenerateENO := "TRUE" } Move(in := 410, out1 => #StateNo)
   END_RUNG
   // the same network as SCL:
   #s410_StWtL1TransBegin := (#s410_StWtL1TransBegin OR #s400_StWtL1S1Down1_T1) AND NOT #sStWtResetRel AND NOT #s410_StWtL1TransBegin_T1;
   IF #s410_StWtL1TransBegin THEN #StateNo := 410; END_IF;
END_REGION

REGION Network 111: Actions for STATE Num:410 StWtL1TransBegin
   RUNG wire#powerrail
      Contact( #s410_StWtL1TransBegin )
      Coil( #qL1TrnsfrConv )
   END_RUNG
   // the same network as SCL:
   #qL1TrnsfrConv := #s410_StWtL1TransBegin;
END_REGION

REGION Network 112: Transition for STATE Num:420 StWtL1TransComplet
   RUNG wire#powerrail
      Contact( #s420_StWtL1TransComplet )
      I_Contact( #sStWtResetRel )
      Contact( #sSst )
      I_Contact( #iAreaClear_TT )
      Contact( #ipalletPrsntAtTT )
      Coil( #s420_StWtL1TransComplet_T1 )
   END_RUNG
   // the same network as SCL:
   #s420_StWtL1TransComplet_T1 := #s420_StWtL1TransComplet AND NOT #sStWtResetRel AND #sSst AND NOT #iAreaClear_TT AND #ipalletPrsntAtTT;
END_REGION

REGION Network 113: STATE Num:420 StWtL1TransComplet
   RUNG wire#powerrail
      Contact( #s420_StWtL1TransComplet )
      wire#w1
      I_Contact( #sStWtResetRel )
      I_Contact( #s420_StWtL1TransComplet_T1 )
      wire#w2
      Coil( #s420_StWtL1TransComplet )
   END_RUNG
   RUNG wire#powerrail
      Contact( #s410_StWtL1TransBegin_T1 )
   END_RUNG wire#w1
   RUNG wire#powerrail
      Contact( #s130_StNextRdyInTransit_1_T2 )
   END_RUNG wire#w1
   RUNG wire#w2
      { S7_GenerateENO := "TRUE" } Move(in := 420, out1 => #StateNo)
   END_RUNG
   // the same network as SCL:
   #s420_StWtL1TransComplet := (#s420_StWtL1TransComplet OR #s410_StWtL1TransBegin_T1 OR #s130_StNextRdyInTransit_1_T2) AND NOT #sStWtResetRel AND NOT #s420_StWtL1TransComplet_T1;
   IF #s420_StWtL1TransComplet THEN #StateNo := 420; END_IF;
END_REGION

REGION Network 114: Transition for STATE Num:430 StNextRdyInTransit_3
   RUNG wire#powerrail
      Contact( #s430_StNextRdyInTransit_3 )
      I_Contact( #sStWtResetRel )
      Contact( #sSst )
      wire#w1
      Contact( #iRTRFrmConv )
      Coil( #s430_StNextRdyInTransit_3_T1 )
   END_RUNG
   RUNG wire#w1
      I_Contact( #s430_StNextRdyInTransit_3_T1 )
      Contact( #iRTRFrmConv )
      Coil( #s430_StNextRdyInTransit_3_T2 )
   END_RUNG
   // the same network as SCL:
   #_w1 := #s430_StNextRdyInTransit_3 AND NOT #sStWtResetRel AND #sSst;
   #s430_StNextRdyInTransit_3_T1 := #_w1 AND #iRTRFrmConv;
   #s430_StNextRdyInTransit_3_T2 := #_w1 AND NOT #s430_StNextRdyInTransit_3_T1 AND #iRTRFrmConv;
END_REGION

REGION Network 115: STATE Num:430 StNextRdyInTransit_3
   RUNG wire#powerrail
      Contact( #s430_StNextRdyInTransit_3 )
      wire#w1
      I_Contact( #sStWtResetRel )
      I_Contact( #s430_StNextRdyInTransit_3_T1 )
      I_Contact( #s430_StNextRdyInTransit_3_T2 )
      wire#w2
      Coil( #s430_StNextRdyInTransit_3 )
   END_RUNG
   RUNG wire#powerrail
      Contact( #s10_StRecovery_T5 )
   END_RUNG wire#w1
   RUNG wire#w2
      { S7_GenerateENO := "TRUE" } Move(in := 430, out1 => #StateNo)
   END_RUNG
   // the same network as SCL:
   #s430_StNextRdyInTransit_3 := (#s430_StNextRdyInTransit_3 OR #s10_StRecovery_T5) AND NOT #sStWtResetRel AND NOT #s430_StNextRdyInTransit_3_T1 AND NOT #s430_StNextRdyInTransit_3_T2;
   IF #s430_StNextRdyInTransit_3 THEN #StateNo := 430; END_IF;
END_REGION
END_FUNCTION_BLOCK
